(* IEC 61131-3 sources: stdmachine/plc/src/04_Objects, 21 files *)

(* ---- FB_AnalogInput.st ---- *)
// Entrée analogique, type 3 (docs/03 § 3.3)
FUNCTION_BLOCK FB_AnalogInput EXTENDS FB_ObjectBase
VAR
    _aSamples : ARRAY[1..100] OF LREAL;
    _nSamples : INT;
    _nNext : INT := 1;
    _fValue : LREAL;                // valeur filtrée, en unité
    _bLowActive : BOOL;
    _bHighActive : BOOL;
END_VAR

METHOD PROTECTED _OnConfigure : BOOL
_nSamples := 0;
_nNext := 1;
_OnConfigure := F_SignalValid(_refCfg.aSignal[1], E_SignalKind.AI) AND _refCfg.aParam[2] <> _refCfg.aParam[1];
END_METHOD

METHOD PROTECTED _OnStart : E_ActStatus
VAR_INPUT
    nAction : UINT;
END_VAR
CASE nAction OF
    GVL_Catalog.AnalogInput_Lire:
        _SetResult(1, _fValue);
        _OnStart := E_ActStatus.Done;
    GVL_Catalog.AnalogInput_AttendreSeuil:
        _OnStart := _OnCycle(nAction);
    GVL_Catalog.AnalogInput_VerifierPlage:
        _SetResult(1, _fValue);
        IF _fValue < _ParamReal(1, -1.0E38) THEN
            _SetJudgement(2, E_Judgement.Low);
        ELSIF _fValue > _ParamReal(2, 1.0E38) THEN
            _SetJudgement(2, E_Judgement.High);
        ELSE
            _SetJudgement(2, E_Judgement.Ok);
        END_IF
        _OnStart := E_ActStatus.Done;
ELSE
    _OnStart := E_ActStatus.Error;
END_CASE
END_METHOD

METHOD PROTECTED _OnCycle : E_ActStatus
VAR_INPUT
    nAction : UINT;
END_VAR
VAR
    bReached : BOOL;
END_VAR
IF _ParamReal(2, 0.0) = 0.0 THEN
    bReached := _fValue >= _ParamReal(1, 0.0);      // au-dessus
ELSE
    bReached := _fValue <= _ParamReal(1, 0.0);      // en dessous
END_IF
IF bReached THEN
    _SetResult(1, _fValue);
    _OnCycle := E_ActStatus.Done;
ELSE
    _OnCycle := E_ActStatus.Busy;
END_IF
END_METHOD

METHOD PROTECTED _ReadHw
_Filter(_Scale(INT_TO_LREAL(F_ReadAI(_refCfg.aSignal[1]))));
END_METHOD

METHOD PROTECTED _Simulate
IF _Forced(1) THEN _Filter(_ForcedValue(1)); END_IF        // valeur forcée en unité
END_METHOD

METHOD PRIVATE _Scale : LREAL
VAR_INPUT
    fRaw : LREAL;
END_VAR
_Scale := _refCfg.aParam[3] + (fRaw - _refCfg.aParam[1]) * (_refCfg.aParam[4] - _refCfg.aParam[3]) / (_refCfg.aParam[2] - _refCfg.aParam[1]);
END_METHOD

METHOD PRIVATE _Filter
VAR_INPUT
    fUnit : LREAL;
END_VAR
VAR
    nWin : INT;
    i : INT;
    fSum : LREAL;
END_VAR
nWin := LIMIT(1, LREAL_TO_INT(_refCfg.aParam[6]), 100);
_aSamples[_nNext] := fUnit;
_nNext := _nNext MOD nWin + 1;
_nSamples := MIN(_nSamples + 1, nWin);
fSum := 0;
FOR i := 1 TO _nSamples DO fSum := fSum + _aSamples[i]; END_FOR
_fValue := fSum / INT_TO_LREAL(_nSamples);
END_METHOD

// Seuils d'alarme : avertissements surveillés en continu, sans mettre l'objet en erreur
METHOD PROTECTED _Monitor
IF _ipAlarms = 0 THEN RETURN; END_IF
IF _fValue < _refCfg.aParam[7] AND NOT _bLowActive THEN
    _ipAlarms.Raise(_stInfo.nGlobalId, GVL_Catalog.AnalogInput_Err100, 0, E_Severity.Warning);
    _bLowActive := TRUE;
ELSIF _fValue >= _refCfg.aParam[7] AND _bLowActive THEN
    _ipAlarms.Clear(_stInfo.nGlobalId, GVL_Catalog.AnalogInput_Err100);
    _bLowActive := FALSE;
END_IF
IF _fValue > _refCfg.aParam[8] AND NOT _bHighActive THEN
    _ipAlarms.Raise(_stInfo.nGlobalId, GVL_Catalog.AnalogInput_Err101, 0, E_Severity.Warning);
    _bHighActive := TRUE;
ELSIF _fValue <= _refCfg.aParam[8] AND _bHighActive THEN
    _ipAlarms.Clear(_stInfo.nGlobalId, GVL_Catalog.AnalogInput_Err101);
    _bHighActive := FALSE;
END_IF
END_METHOD

METHOD PROTECTED _Publish
_stStatus.aValue[1] := _fValue;
END_METHOD

PROPERTY Value : LREAL
GET
Value := _fValue;
END_GET
END_PROPERTY
END_FUNCTION_BLOCK

(* ---- FB_AnalogOutput.st ---- *)
// Sortie analogique, type 4 (docs/03 § 3.4)
FUNCTION_BLOCK FB_AnalogOutput EXTENDS FB_ObjectBase
VAR
    _fValue : LREAL;                // valeur commandée, en unité
    _fStart : LREAL;
    _fTarget : LREAL;
    _fRampMs : LREAL;
    _fElapsed : LREAL;
END_VAR

METHOD PROTECTED _OnConfigure : BOOL
_OnConfigure := F_SignalValid(_refCfg.aSignal[1], E_SignalKind.AO) AND _refCfg.aParam[4] <> _refCfg.aParam[3];
END_METHOD

METHOD PROTECTED _DefaultTimeoutMs : UDINT
VAR_INPUT
    nAction : UINT;
END_VAR
IF nAction = GVL_Catalog.AnalogOutput_EcrireAvecRampe THEN
    _DefaultTimeoutMs := LREAL_TO_UDINT(MAX(_ParamReal(2, 0.0), 0.0)) + 1000;
ELSE
    _DefaultTimeoutMs := 0;
END_IF
END_METHOD

METHOD PROTECTED _OnStart : E_ActStatus
VAR_INPUT
    nAction : UINT;
END_VAR
_fStart := _fValue;
_fElapsed := 0;
CASE nAction OF
    GVL_Catalog.AnalogOutput_Ecrire:
        _fTarget := _Limit(_ParamReal(1, _fValue));
        _fRampMs := 0;
    GVL_Catalog.AnalogOutput_EcrireAvecRampe:
        _fTarget := _Limit(_ParamReal(1, _fValue));
        _fRampMs := MAX(_ParamReal(2, 0.0), 0.0);
    GVL_Catalog.AnalogOutput_ValeurSure:
        _fTarget := _Limit(_refCfg.aParam[8]);
        _fRampMs := 0;
ELSE
    _OnStart := E_ActStatus.Error;
    RETURN;
END_CASE
_OnStart := _OnCycle(nAction);
END_METHOD

METHOD PROTECTED _OnCycle : E_ActStatus
VAR_INPUT
    nAction : UINT;
END_VAR
VAR
    fNext : LREAL;
    fMaxStep : LREAL;
END_VAR
_fElapsed := _fElapsed + F_CycleMs();
IF _fRampMs > 0 THEN
    fNext := _fStart + (_fTarget - _fStart) * MIN(1.0, _fElapsed / _fRampMs);
ELSE
    fNext := _fTarget;
END_IF
// Variation maximale P9 (unité/s), 0 = illimitée
IF _refCfg.aParam[9] > 0 THEN
    fMaxStep := _refCfg.aParam[9] * F_CycleMs() / 1000.0;
    fNext := LIMIT(_fValue - fMaxStep, fNext, _fValue + fMaxStep);
END_IF
_fValue := fNext;
IF ABS(_fValue - _fTarget) < 1.0E-9 THEN _OnCycle := E_ActStatus.Done; ELSE _OnCycle := E_ActStatus.Busy; END_IF
END_METHOD

METHOD PRIVATE _Limit : LREAL
VAR_INPUT
    fValue : LREAL;
END_VAR
_Limit := LIMIT(_refCfg.aParam[6], fValue, _refCfg.aParam[7]);
END_METHOD

METHOD PROTECTED _SafeState
_fValue := _Limit(_refCfg.aParam[8]);
END_METHOD

METHOD PROTECTED _WriteHw
VAR
    fRaw : LREAL;
END_VAR
fRaw := _refCfg.aParam[1] + (_fValue - _refCfg.aParam[3]) * (_refCfg.aParam[2] - _refCfg.aParam[1]) / (_refCfg.aParam[4] - _refCfg.aParam[3]);
F_WriteAO(_refCfg.aSignal[1], LREAL_TO_INT(LIMIT(-32768.0, fRaw, 32767.0)));
END_METHOD

METHOD PROTECTED _Publish
_stStatus.aValue[1] := _fValue;
END_METHOD
END_FUNCTION_BLOCK

(* ---- FB_Axis.st ---- *)
// Axe linéaire (type 11) et axe rotatif (type 12), docs/03 § 4.2 et docs/04 § 12.
// Matériel : D = n° de l'axe dans GVL_Hw.aAxis (pointeur donné par GVL_IoRef). Blocs Tc2_MC2.
// L'override effectif est appliqué par MC_Power.Override : il ralentit le mouvement en cours sans le relancer.
FUNCTION_BLOCK FB_Axis EXTENDS FB_ObjectBase
VAR
    _pAxis : POINTER TO AXIS_REF;
    _bRotary : BOOL;
    _fbPower : MC_Power;
    _fbReset : MC_Reset;
    _fbHome : MC_Home;
    _fbMoveAbs : MC_MoveAbsolute;
    _fbMoveMod : MC_MoveModulo;
    _fbMoveRel : MC_MoveRelative;
    _fbHalt : MC_Halt;
    _fbStop : MC_Stop;
    _fbJog : MC_Jog;
    _bEnable : BOOL;                // alimentation demandée
    _bPowered : BOOL;
    _bWasPowered : BOOL;
    _bHomed : BOOL;
    _fActPos : LREAL;
    _fActVel : LREAL;
    _fTarget : LREAL;
    _fStartPos : LREAL;
    _fVelo : LREAL;
    _fAcc : LREAL;
    _fDec : LREAL;
    _nDirection : INT;              // rotatif : 0 plus court, 1 positif, 2 négatif
    _bExecute : BOOL;               // front de commande de l'action en cours
    _bStopping : BOOL;              // Abort : arrêt en cours
    _fOverride : LREAL := 100.0;
    // Simulation : profil trapézoïdal
    _fSimPos : LREAL;
    _fSimVel : LREAL;
    _fSimInitMs : LREAL;
    _nJogDir : INT;                 // +1, -1, 0
END_VAR

METHOD PROTECTED _OnConfigure : BOOL
_bRotary := _refCfg.nType = GVL_Catalog.Type_RotaryAxis;
_pAxis := F_AxisRef(_refCfg.nDevice);
_bEnable := FALSE;
_bHomed := FALSE;
_fSimVel := 0;
_OnConfigure := _pAxis <> 0 OR _IsSimulated();
END_METHOD

METHOD PROTECTED _NeedsInit : BOOL
_NeedsInit := TRUE;
END_METHOD

METHOD PROTECTED _IsAllowedNotInit : BOOL
VAR_INPUT
    nAction : UINT;
END_VAR
_IsAllowedNotInit := nAction = GVL_Catalog.LinearAxis_PowerOn OR nAction = GVL_Catalog.LinearAxis_PowerOff
                     OR nAction = GVL_Catalog.LinearAxis_Init OR nAction = GVL_Catalog.LinearAxis_AcquitterErreur
                     OR nAction = GVL_Catalog.LinearAxis_LirePosition
                     OR nAction = GVL_Catalog.LinearAxis_JogPlus OR nAction = GVL_Catalog.LinearAxis_JogMoins;
END_METHOD

METHOD PROTECTED _ManualOverride : LREAL
_ManualOverride := LIMIT(0.0, _refCfg.aParam[12], 100.0);
END_METHOD

METHOD PROTECTED _DefaultTimeoutMs : UDINT
VAR_INPUT
    nAction : UINT;
END_VAR
VAR
    fDist : LREAL;
END_VAR
// Move absolu et relatif : 2 × (distance ÷ vitesse + vitesse ÷ accélération) × 1000 + 1000 ms, à 100 %
IF nAction = GVL_Catalog.LinearAxis_MoveAbsolu OR nAction = GVL_Catalog.LinearAxis_MoveRelatif THEN
    IF nAction = GVL_Catalog.LinearAxis_MoveAbsolu THEN fDist := ABS(_TargetOf() - _fActPos); ELSE fDist := ABS(_ParamReal(1, 0.0)); END_IF
    _Kinematics();
    IF _fVelo > 0 AND _fAcc > 0 THEN
        _DefaultTimeoutMs := LREAL_TO_UDINT(2.0 * (fDist / _fVelo + _fVelo / _fAcc) * 1000.0 + 1000.0);
    ELSE
        _DefaultTimeoutMs := 30000;
    END_IF
ELSE
    _DefaultTimeoutMs := SUPER^._DefaultTimeoutMs(nAction);
END_IF
END_METHOD

METHOD PRIVATE _TargetOf : LREAL
// Une position nommée : composante P13 (X, Y, Z) ou C pour un rotatif, plus le décalage (hauteur d'approche)
IF _stParams.aKind[1] = E_ParamKind.Position THEN
    IF _bRotary THEN
        _TargetOf := _stParams.stPos.fC;
    ELSE
        CASE LREAL_TO_INT(_refCfg.aParam[13]) OF
            1: _TargetOf := _stParams.stPos.fY;
            2: _TargetOf := _stParams.stPos.fZ;
        ELSE
            _TargetOf := _stParams.stPos.fX;
        END_CASE
    END_IF
    _TargetOf := _TargetOf + _stParams.aReal[1];
ELSE
    _TargetOf := _stParams.aReal[1];
END_IF
END_METHOD

METHOD PRIVATE _Kinematics
VAR
    fAccPct : LREAL;
END_VAR
_fVelo := MAX(_refCfg.aParam[1], 0.001) * F_ParamSpeed(_stParams, 2, _refCfg, 2) / 100.0;
fAccPct := LIMIT(1.0, _ParamReal(3, 100.0), 100.0);
IF _stParams.aKind[3] = E_ParamKind.Unused THEN fAccPct := 100.0; END_IF
_fAcc := MAX(_refCfg.aParam[2], 0.001) * fAccPct / 100.0;
_fDec := MAX(_refCfg.aParam[3], 0.001) * fAccPct / 100.0;
END_METHOD

METHOD PROTECTED _OnStart : E_ActStatus
VAR_INPUT
    nAction : UINT;
END_VAR
_bExecute := FALSE;
_bStopping := FALSE;
_fStartPos := _fActPos;
CASE nAction OF
    GVL_Catalog.LinearAxis_PowerOn:
        _bEnable := TRUE;
        _OnStart := E_ActStatus.Busy;
    GVL_Catalog.LinearAxis_PowerOff:
        _bEnable := FALSE;
        _OnStart := E_ActStatus.Busy;
    GVL_Catalog.LinearAxis_Init:
        IF NOT _bPowered THEN _Fail(GVL_Catalog.LinearAxis_Err105, 0); _OnStart := E_ActStatus.Error; RETURN; END_IF
        _bHomed := FALSE;
        _bInitialized := FALSE;
        _fSimInitMs := 0;
        _OnStart := E_ActStatus.Busy;
    GVL_Catalog.LinearAxis_MoveAbsolu, GVL_Catalog.LinearAxis_MoveRelatif:
        IF NOT _bPowered THEN _Fail(GVL_Catalog.LinearAxis_Err105, 0); _OnStart := E_ActStatus.Error; RETURN; END_IF
        IF NOT _bHomed THEN _Fail(GVL_Catalog.LinearAxis_Err100, 0); _OnStart := E_ActStatus.Error; RETURN; END_IF
        IF nAction = GVL_Catalog.LinearAxis_MoveAbsolu THEN
            _fTarget := _TargetOf();
            _nDirection := LREAL_TO_INT(_ParamReal(4, _refCfg.aParam[14]));
        ELSE
            _fTarget := _fActPos + _ParamReal(1, 0.0);
        END_IF
        IF _refCfg.aParam[7] = 1 AND (_fTarget < _refCfg.aParam[5] OR _fTarget > _refCfg.aParam[6]) THEN
            _Fail(GVL_Catalog.LinearAxis_Err101, 0);
            _OnStart := E_ActStatus.Error;
            RETURN;
        END_IF
        _Kinematics();
        _OnStart := E_ActStatus.Busy;
    GVL_Catalog.LinearAxis_Stop:
        _OnStart := E_ActStatus.Busy;
    GVL_Catalog.LinearAxis_AcquitterErreur:
        _OnStart := E_ActStatus.Busy;
    GVL_Catalog.LinearAxis_LirePosition:
        _SetResult(1, _fActPos);
        _OnStart := E_ActStatus.Done;
    GVL_Catalog.LinearAxis_JogPlus, GVL_Catalog.LinearAxis_JogMoins:
        IF NOT _bPowered THEN _Fail(GVL_Catalog.LinearAxis_Err105, 0); _OnStart := E_ActStatus.Error; RETURN; END_IF
        _fVelo := MAX(_refCfg.aParam[1], 0.001) * F_ParamSpeed(_stParams, 1, _refCfg, 1) / 100.0;
        IF NOT _bHomed THEN _fVelo := MAX(_refCfg.aParam[1], 0.001) * F_ParamSpeed(_stParams, 0, _refCfg, 1) / 100.0; END_IF   // V1 imposée
        _fAcc := MAX(_refCfg.aParam[2], 0.001);
        _fDec := MAX(_refCfg.aParam[3], 0.001);
        _nJogDir := SEL(nAction = GVL_Catalog.LinearAxis_JogPlus, -1, 1);
        _OnStart := E_ActStatus.Busy;       // le jog dure jusqu'à Abort (canal manuel, docs/05 § 7)
ELSE
    _OnStart := E_ActStatus.Error;
END_CASE
END_METHOD

METHOD PROTECTED _OnCycle : E_ActStatus
VAR_INPUT
    nAction : UINT;
END_VAR
_OnCycle := E_ActStatus.Busy;
CASE nAction OF
    GVL_Catalog.LinearAxis_PowerOn:
        IF _bPowered THEN _OnCycle := E_ActStatus.Done; END_IF
    GVL_Catalog.LinearAxis_PowerOff:
        IF NOT _bPowered THEN _OnCycle := E_ActStatus.Done; END_IF
    GVL_Catalog.LinearAxis_Init:
        IF _IsSimulated() THEN
            _fSimInitMs := _fSimInitMs + F_CycleMs();
            IF _fSimInitMs >= 1500.0 THEN
                _fSimPos := _refCfg.aParam[8];
                _fSimVel := 0;
                _bHomed := TRUE;
            END_IF
        ELSE
            _bExecute := TRUE;
            IF _fbHome.Done THEN _bHomed := TRUE; END_IF
            IF _fbHome.Error THEN _Fail(GVL_Catalog.LinearAxis_Err102, _fbHome.ErrorID); _OnCycle := E_ActStatus.Error; RETURN; END_IF
        END_IF
        IF _bHomed THEN
            _bInitialized := TRUE;
            _bExecute := FALSE;
            _OnCycle := E_ActStatus.Done;
        END_IF
    GVL_Catalog.LinearAxis_MoveAbsolu, GVL_Catalog.LinearAxis_MoveRelatif:
        IF _IsSimulated() THEN
            IF ABS(_fSimPos - _fTarget) <= MAX(_refCfg.aParam[4], 1.0E-6) AND ABS(_fSimVel) < 1.0E-6 THEN _OnCycle := E_ActStatus.Done; END_IF
        ELSE
            _bExecute := TRUE;
            IF _fbMoveAbs.Done OR _fbMoveRel.Done OR _fbMoveMod.Done THEN _OnCycle := E_ActStatus.Done; END_IF
            IF _fbMoveAbs.Error OR _fbMoveRel.Error OR _fbMoveMod.Error THEN
                _Fail(GVL_Catalog.LinearAxis_Err102, _fbMoveAbs.ErrorID OR _fbMoveRel.ErrorID OR _fbMoveMod.ErrorID);
                _OnCycle := E_ActStatus.Error;
                RETURN;
            END_IF
        END_IF
        IF _OnCycle = E_ActStatus.Done THEN
            _bExecute := FALSE;
            _SetResult(1, _fActPos);
        END_IF
    GVL_Catalog.LinearAxis_Stop:
        IF _IsSimulated() THEN
            IF ABS(_fSimVel) < 1.0E-6 THEN _OnCycle := E_ActStatus.Done; END_IF
        ELSE
            _bExecute := TRUE;
            IF _fbHalt.Done THEN _bExecute := FALSE; _OnCycle := E_ActStatus.Done; END_IF
        END_IF
    GVL_Catalog.LinearAxis_AcquitterErreur:
        IF _IsSimulated() THEN
            _OnCycle := E_ActStatus.Done;
        ELSE
            _bExecute := TRUE;
            IF _fbReset.Done OR _fbReset.Error THEN _bExecute := FALSE; _OnCycle := E_ActStatus.Done; END_IF
        END_IF
    GVL_Catalog.LinearAxis_JogPlus, GVL_Catalog.LinearAxis_JogMoins:
        ;                               // jusqu'à Abort
END_CASE
_CallMotion();
END_METHOD

METHOD PROTECTED _OnAbort
VAR_INPUT
    nAction : UINT;
END_VAR
// Arrêt avec la décélération maximale, puis P11 (0 alimentation maintenue, 1 coupée)
_bExecute := FALSE;
_nJogDir := 0;
_bStopping := TRUE;
END_METHOD

METHOD PROTECTED _SafeState
IF _refCfg.aParam[11] = 1 THEN _bEnable := FALSE; END_IF
END_METHOD

METHOD PROTECTED _OnAck : BOOL
IF _IsSimulated() OR _pAxis = 0 THEN
    _OnAck := TRUE;
    RETURN;
END_IF
_fbReset(Axis := _pAxis^, Execute := TRUE);
IF _fbReset.Done OR _fbReset.Error THEN
    _fbReset(Axis := _pAxis^, Execute := FALSE);
    _OnAck := TRUE;
END_IF
END_METHOD

METHOD PROTECTED _ApplyOverride
VAR_INPUT
    fPercent : LREAL;
END_VAR
_fOverride := LIMIT(0.0, fPercent, 100.0);
END_METHOD

METHOD PROTECTED _ReadHw
IF _pAxis = 0 THEN RETURN; END_IF
_pAxis^.ReadStatus();
_fActPos := _pAxis^.NcToPlc.ActPos;
_fActVel := _pAxis^.NcToPlc.ActVelo;
_bHomed := _bHomed OR _pAxis^.Status.Homed;
_fbPower(Axis := _pAxis^, Enable := _bEnable, Enable_Positive := _bEnable, Enable_Negative := _bEnable, Override := _fOverride);
_bPowered := _fbPower.Status;
IF NOT _bExecute AND _eState <> E_ObjState.Busy THEN _CallMotion(); END_IF    // remet les Execute à FALSE
END_METHOD

METHOD PRIVATE _CallMotion
VAR
    bAbs : BOOL;
    bRel : BOOL;
    bMod : BOOL;
    eDir : MC_Direction;
END_VAR
IF _IsSimulated() OR _pAxis = 0 THEN RETURN; END_IF
bAbs := _bExecute AND _nAction = GVL_Catalog.LinearAxis_MoveAbsolu AND NOT (_bRotary AND _refCfg.aParam[7] = 0);
bMod := _bExecute AND _nAction = GVL_Catalog.LinearAxis_MoveAbsolu AND _bRotary AND _refCfg.aParam[7] = 0;
bRel := _bExecute AND _nAction = GVL_Catalog.LinearAxis_MoveRelatif;
CASE _nDirection OF
    1: eDir := MC_Positive_Direction;
    2: eDir := MC_Negative_Direction;
ELSE
    eDir := MC_Shortest_Way;
END_CASE
_fbHome(Axis := _pAxis^, Execute := _bExecute AND _nAction = GVL_Catalog.LinearAxis_Init, Position := _refCfg.aParam[8],
        HomingMode := SEL(LREAL_TO_INT(_refCfg.aParam[9]) = 3, MC_DefaultHoming, MC_Direct));
_fbMoveAbs(Axis := _pAxis^, Execute := bAbs, Position := _fTarget, Velocity := _fVelo, Acceleration := _fAcc, Deceleration := _fDec);
_fbMoveMod(Axis := _pAxis^, Execute := bMod, Position := _fTarget, Velocity := _fVelo, Acceleration := _fAcc, Deceleration := _fDec, Direction := eDir);
_fbMoveRel(Axis := _pAxis^, Execute := bRel, Distance := _fTarget - _fStartPos, Velocity := _fVelo, Acceleration := _fAcc, Deceleration := _fDec);
_fbHalt(Axis := _pAxis^, Execute := _bExecute AND _nAction = GVL_Catalog.LinearAxis_Stop);
_fbReset(Axis := _pAxis^, Execute := _bExecute AND _nAction = GVL_Catalog.LinearAxis_AcquitterErreur);
_fbJog(Axis := _pAxis^, JogForward := _nJogDir > 0, JogBackwards := _nJogDir < 0, Mode := MC_JOGMODE_CONTINOUS,
       Velocity := _fVelo, Acceleration := _fAcc, Deceleration := _fDec);
_fbStop(Axis := _pAxis^, Execute := _bStopping);
IF _bStopping AND (_fbStop.Done OR _fbStop.Error) THEN
    _bStopping := FALSE;
    _fbStop(Axis := _pAxis^, Execute := FALSE);
END_IF
END_METHOD

METHOD PROTECTED _Monitor
IF _IsSimulated() OR _pAxis = 0 THEN
    _bWasPowered := _bPowered;
    RETURN;
END_IF
IF _pAxis^.Status.Error AND _eState <> E_ObjState.Error THEN
    IF _pAxis^.Status.ErrorID = 16#4550 OR _pAxis^.Status.ErrorID = 16#4551 THEN
        _Fail(GVL_Catalog.LinearAxis_Err103, _pAxis^.Status.ErrorID);      // erreur de suivi
    ELSE
        _Fail(GVL_Catalog.LinearAxis_Err102, _pAxis^.Status.ErrorID);      // erreur du drive (sous-code NC)
    END_IF
ELSIF _bWasPowered AND NOT _bPowered AND _bEnable AND _eState <> E_ObjState.Error THEN
    _Fail(GVL_Catalog.LinearAxis_Err104, 0);                                 // perte d'alimentation
END_IF
_bWasPowered := _bPowered;
END_METHOD

METHOD PROTECTED _Simulate
VAR
    fDt : LREAL;
    fVmax : LREAL;
    fDist : LREAL;
    fBrake : LREAL;
    fDir : LREAL;
END_VAR
fDt := F_CycleMs() / 1000.0;
_bPowered := _bEnable;
fVmax := _fVelo * _fOverride / 100.0;
IF _bStopping THEN
    // arrêt avec la décélération maximale
    IF _fSimVel > 0 THEN _fSimVel := MAX(0.0, _fSimVel - _refCfg.aParam[3] * fDt); ELSE _fSimVel := MIN(0.0, _fSimVel + _refCfg.aParam[3] * fDt); END_IF
    IF ABS(_fSimVel) < 1.0E-9 THEN _bStopping := FALSE; END_IF
ELSIF _eState = E_ObjState.Busy AND (_nAction = GVL_Catalog.LinearAxis_JogPlus OR _nAction = GVL_Catalog.LinearAxis_JogMoins) THEN
    _fSimVel := LIMIT(-fVmax, _fSimVel + INT_TO_LREAL(_nJogDir) * _fAcc * fDt, fVmax);
ELSIF _eState = E_ObjState.Busy AND (_nAction = GVL_Catalog.LinearAxis_MoveAbsolu OR _nAction = GVL_Catalog.LinearAxis_MoveRelatif) THEN
    fDist := _fTarget - _fSimPos;
    fDir := SEL(fDist >= 0, -1.0, 1.0);
    fBrake := _fSimVel * _fSimVel / (2.0 * MAX(_fDec, 0.001));
    IF ABS(fDist) <= fBrake THEN
        _fSimVel := _fSimVel - fDir * _fDec * fDt;          // décélération
        IF fDir * _fSimVel < 0 THEN _fSimVel := 0; END_IF
    ELSE
        _fSimVel := LIMIT(-fVmax, _fSimVel + fDir * _fAcc * fDt, fVmax);
    END_IF
    IF ABS(fDist) <= ABS(_fSimVel * fDt) OR (ABS(_fSimVel) < 1.0E-9 AND ABS(fDist) <= MAX(_refCfg.aParam[4], 1.0E-6)) THEN
        _fSimPos := _fTarget;
        _fSimVel := 0;
    END_IF
ELSIF _eState = E_ObjState.Busy AND _nAction = GVL_Catalog.LinearAxis_Stop THEN
    IF _fSimVel > 0 THEN _fSimVel := MAX(0.0, _fSimVel - _fDec * fDt); ELSE _fSimVel := MIN(0.0, _fSimVel + _fDec * fDt); END_IF
ELSE
    _fSimVel := 0;
END_IF
_fSimPos := _fSimPos + _fSimVel * fDt;
_fActPos := _fSimPos;
_fActVel := _fSimVel;
END_METHOD

METHOD PROTECTED _Publish
_stStatus.aValue[1] := _fActPos;
_stStatus.aValue[2] := _fActVel;
_stStatus.aValue[3] := BOOL_TO_LREAL(_bPowered);
_stStatus.aValue[4] := BOOL_TO_LREAL(_bHomed);
IF _eState = E_ObjState.Busy AND ABS(_fTarget - _fStartPos) > 1.0E-9
   AND (_nAction = GVL_Catalog.LinearAxis_MoveAbsolu OR _nAction = GVL_Catalog.LinearAxis_MoveRelatif) THEN
    _stStatus.fProgress := LREAL_TO_REAL(LIMIT(0.0, ABS(_fActPos - _fStartPos) / ABS(_fTarget - _fStartPos), 1.0));
END_IF
END_METHOD

PROPERTY ActualPosition : LREAL
GET
ActualPosition := _fActPos;
END_GET
END_PROPERTY
END_FUNCTION_BLOCK

(* ---- FB_Beacon.st ---- *)
// Balise, type 50 (docs/03 § 8.1) : pilotée par le séquenceur ; actions de test en manuel seulement
FUNCTION_BLOCK FB_Beacon EXTENDS FB_ObjectBase IMPLEMENTS I_Beacon
VAR
    _nPattern : UINT;
    _bBuzzerReq : BOOL;
    _fBlink : LREAL;
    _bPhase : BOOL;
    _nTestColor : INT := -1;        // test manuel : 0 rouge, 1 orange, 2 vert, 3 bleu, 4 buzzer
    _fTestMs : LREAL;
    _fBuzzMs : LREAL;               // durée de buzzer demandée (0 = jusqu'à acquittement)
    _fBuzzElapsed : LREAL;
    _aOut : ARRAY[1..5] OF BOOL;    // rouge, orange, vert, bleu, buzzer
END_VAR

METHOD SetPattern
VAR_INPUT
    nPattern : UINT;
    bBuzzer : BOOL;
END_VAR
IF bBuzzer AND NOT _bBuzzerReq THEN _fBuzzElapsed := 0; END_IF
_nPattern := nPattern;
_bBuzzerReq := bBuzzer;
END_METHOD

METHOD PROTECTED _OnStart : E_ActStatus
VAR_INPUT
    nAction : UINT;
END_VAR
_fBuzzElapsed := 0;
CASE nAction OF
    GVL_Catalog.Beacon_Tester:
        _nTestColor := LIMIT(0, LREAL_TO_INT(_ParamReal(1, 0.0)), 4);
        _fTestMs := MAX(_ParamReal(2, 2000.0), 100.0);
        _OnStart := E_ActStatus.Busy;
    GVL_Catalog.Beacon_Buzzer:
        _nTestColor := 4;
        _fTestMs := MAX(_ParamReal(1, 1000.0), 100.0);
        _OnStart := E_ActStatus.Busy;
ELSE
    _OnStart := E_ActStatus.Error;
END_CASE
END_METHOD

METHOD PROTECTED _OnCycle : E_ActStatus
VAR_INPUT
    nAction : UINT;
END_VAR
IF _fElapsedMs >= _fTestMs THEN
    _nTestColor := -1;
    _OnCycle := E_ActStatus.Done;
ELSE
    _OnCycle := E_ActStatus.Busy;
END_IF
END_METHOD

METHOD PROTECTED _OnAbort
VAR_INPUT
    nAction : UINT;
END_VAR
_nTestColor := -1;
END_METHOD

METHOD PROTECTED _Monitor
VAR
    fPeriod : LREAL;
    i : INT;
END_VAR
fPeriod := MAX(_refCfg.aParam[1], 100.0);
_fBlink := _fBlink + F_CycleMs();
IF _fBlink >= fPeriod / 2.0 THEN
    _fBlink := 0;
    _bPhase := NOT _bPhase;
END_IF
FOR i := 1 TO 5 DO _aOut[i] := FALSE; END_FOR
IF _nTestColor >= 0 THEN
    _aOut[_nTestColor + 1] := TRUE;
    RETURN;
END_IF
_aOut[1] := (_nPattern AND GVL_BeaconBits.RED) <> 0 OR ((_nPattern AND GVL_BeaconBits.RED_BLINK) <> 0 AND _bPhase);
_aOut[2] := (_nPattern AND GVL_BeaconBits.ORANGE) <> 0 OR ((_nPattern AND GVL_BeaconBits.ORANGE_BLINK) <> 0 AND _bPhase);
_aOut[3] := (_nPattern AND GVL_BeaconBits.GREEN) <> 0 OR ((_nPattern AND GVL_BeaconBits.GREEN_BLINK) <> 0 AND _bPhase);
_aOut[4] := (_nPattern AND GVL_BeaconBits.BLUE) <> 0 OR ((_nPattern AND GVL_BeaconBits.BLUE_BLINK) <> 0 AND _bPhase);
IF _bBuzzerReq THEN
    _fBuzzElapsed := _fBuzzElapsed + F_CycleMs();
    _aOut[5] := _refCfg.aParam[2] <= 0 OR _fBuzzElapsed < _refCfg.aParam[2];
END_IF
END_METHOD

METHOD PROTECTED _WriteHw
VAR
    i : USINT;
END_VAR
FOR i := 1 TO 5 DO F_WriteDO(_refCfg.aSignal[i], _aOut[i]); END_FOR
END_METHOD

METHOD PROTECTED _Publish
VAR
    i : INT;
    nBits : DWORD;
END_VAR
FOR i := 1 TO 5 DO
    IF _aOut[i] THEN nBits := nBits OR SHL(DWORD#1, i - 1); END_IF
END_FOR
_stStatus.aValue[1] := DWORD_TO_LREAL(nBits);
END_METHOD
END_FUNCTION_BLOCK

(* ---- FB_Counter.st ---- *)
// Compteur, type 53 (docs/03 § 8.4)
FUNCTION_BLOCK FB_Counter EXTENDS FB_ObjectBase IMPLEMENTS I_OrderAware
VAR
    _bStarted : BOOL;               // faux au démarrage du PLC (P4 = 0 : la valeur repart de P1)
END_VAR
VAR PERSISTENT
    _fValue : LREAL;
END_VAR

METHOD PROTECTED _OnConfigure : BOOL
IF _bNewObject THEN _fValue := _refCfg.aParam[1]; END_IF
_OnConfigure := TRUE;
END_METHOD

METHOD PROTECTED _OnStart : E_ActStatus
VAR_INPUT
    nAction : UINT;
END_VAR
CASE nAction OF
    GVL_Catalog.Counter_Incrementer:
        _fValue := _fValue + _ParamReal(1, 1.0);
        _SetResult(1, _fValue);
        IF _refCfg.aParam[2] > 0 AND _fValue > _refCfg.aParam[2] THEN
            _Fail(GVL_Catalog.Counter_Err100, LREAL_TO_UDINT(_fValue));
            _OnStart := E_ActStatus.Error;
            RETURN;
        END_IF
    GVL_Catalog.Counter_Lire:
        _SetResult(1, _fValue);
    GVL_Catalog.Counter_RemettreAZero:
        _fValue := _refCfg.aParam[1];
    GVL_Catalog.Counter_Comparer:
        _SetResult(1, BOOL_TO_LREAL(_fValue >= _ParamReal(1, 0.0)));
ELSE
    _OnStart := E_ActStatus.Error;
    RETURN;
END_CASE
_OnStart := E_ActStatus.Done;
END_METHOD

// Remise à zéro au changement d'OF (P3), appelée par le séquenceur général
METHOD OnOrderChange
IF _refCfg.aParam[3] = 1 THEN _fValue := _refCfg.aParam[1]; END_IF
END_METHOD

METHOD PROTECTED _Monitor
IF NOT _bStarted THEN
    _bStarted := TRUE;
    IF _refCfg.aParam[4] = 0 THEN _fValue := _refCfg.aParam[1]; END_IF
END_IF
END_METHOD

METHOD PROTECTED _Publish
_stStatus.aValue[1] := _fValue;
END_METHOD
END_FUNCTION_BLOCK

(* ---- FB_Cylinder.st ---- *)
// Vérin, type 10 (docs/03 § 4.1, exemple complet de docs/04 § 11)
FUNCTION_BLOCK FB_Cylinder EXTENDS FB_ObjectBase
VAR
    _bBistable : BOOL;
    _tSettleMs : LREAL;
    _tNoSensorMs : LREAL;
    _eSafe : USINT;                 // 0 Repos, 1 Travail, 2 Maintien
    _bCmdWork : BOOL;               // sortie travail commandée
    _bAtWork : BOOL;                // capteurs (lus ou simulés)
    _bAtRest : BOOL;
    _bHasWorkSensor : BOOL;
    _bHasRestSensor : BOOL;
    _fSettle : LREAL;
    _fMove : LREAL;
    _fSimPos : LREAL;               // simulation : 0 = repos, 1 = travail
    _nReached : USINT;              // 0 aucune, 1 repos, 2 travail : dernière position atteinte par une action
END_VAR

METHOD PROTECTED _OnConfigure : BOOL
_bBistable := _refCfg.aParam[1] = 1;
_tSettleMs := LIMIT(0.0, _refCfg.aParam[2], 5000.0);
_tNoSensorMs := MAX(_refCfg.aParam[3], 10.0);
_eSafe := LREAL_TO_USINT(_refCfg.aParam[4]);
_bHasWorkSensor := F_SignalValid(_refCfg.aSignal[3], E_SignalKind.DI);
_bHasRestSensor := F_SignalValid(_refCfg.aSignal[4], E_SignalKind.DI);
_nReached := 0;
_OnConfigure := F_SignalValid(_refCfg.aSignal[1], E_SignalKind.DO)
                AND (NOT _bBistable OR F_SignalValid(_refCfg.aSignal[2], E_SignalKind.DO));
END_METHOD

METHOD PROTECTED _DefaultTimeoutMs : UDINT
VAR_INPUT
    nAction : UINT;
END_VAR
_DefaultTimeoutMs := SEL(_bHasWorkSensor OR _bHasRestSensor, LREAL_TO_UDINT(_tNoSensorMs) + 500, 2000);
END_METHOD

METHOD PROTECTED _OnStart : E_ActStatus
VAR_INPUT
    nAction : UINT;
END_VAR
CASE nAction OF
    GVL_Catalog.Cylinder_MoveTravail, GVL_Catalog.Cylinder_MoveRepos:
        _fMove := 0;
        _fSettle := 0;
        _nReached := 0;
        _OnStart := E_ActStatus.Busy;   // la commande est posée dans _OnCycle (attente si override 0 %)
    GVL_Catalog.Cylinder_LirePosition:
        _SetResult(1, _PositionCode());
        _OnStart := E_ActStatus.Done;
ELSE
    _OnStart := E_ActStatus.Error;
END_CASE
END_METHOD

METHOD PROTECTED _OnCycle : E_ActStatus
VAR_INPUT
    nAction : UINT;
END_VAR
VAR
    bTarget : BOOL;
    bSensorOk : BOOL;
    fCycleMs : LREAL;
END_VAR
fCycleMs := F_CycleMs();
IF _fEffOverride <= 0 AND _fMove = 0 THEN _OnCycle := E_ActStatus.Busy; RETURN; END_IF   // 0 % : on attend
bTarget := nAction = GVL_Catalog.Cylinder_MoveTravail;
_bCmdWork := bTarget;
_fMove := _fMove + fCycleMs;
// Capteur de départ toujours actif après 500 ms : vérin bloqué (erreur 102)
IF _fMove >= 500.0 AND ((bTarget AND _bHasRestSensor AND _bAtRest) OR (NOT bTarget AND _bHasWorkSensor AND _bAtWork)) THEN
    _Fail(GVL_Catalog.Cylinder_Err102, 0);
    _OnCycle := E_ActStatus.Error;
    RETURN;
END_IF
IF bTarget THEN
    bSensorOk := SEL(_bHasWorkSensor, _fMove >= _tNoSensorMs, _bAtWork AND NOT _bAtRest);
ELSE
    bSensorOk := SEL(_bHasRestSensor, _fMove >= _tNoSensorMs, _bAtRest AND NOT _bAtWork);
END_IF
IF bSensorOk THEN _fSettle := _fSettle + fCycleMs; ELSE _fSettle := 0; END_IF
IF _fSettle >= _tSettleMs THEN
    _nReached := SEL(bTarget, 1, 2);
    _OnCycle := E_ActStatus.Done;
ELSE
    _OnCycle := E_ActStatus.Busy;
END_IF
END_METHOD

METHOD PROTECTED _SafeState
CASE _eSafe OF
    0: _bCmdWork := FALSE;
    1: _bCmdWork := TRUE;
END_CASE                            // 2 : maintien
END_METHOD

METHOD PROTECTED _Monitor
IF _bAtWork AND _bAtRest THEN
    IF _eState <> E_ObjState.Error THEN _Fail(GVL_Catalog.Cylinder_Err100, 0); END_IF
ELSIF _eState = E_ObjState.Ready THEN
    // Perte du capteur de la position atteinte hors mouvement (erreur 101)
    IF (_nReached = 2 AND _bHasWorkSensor AND NOT _bAtWork) OR (_nReached = 1 AND _bHasRestSensor AND NOT _bAtRest) THEN
        _Fail(GVL_Catalog.Cylinder_Err101, _nReached);
        _nReached := 0;
    END_IF
END_IF
END_METHOD

METHOD PROTECTED _ReadHw
_bAtWork := F_ReadDI(_refCfg.aSignal[3]);
_bAtRest := F_ReadDI(_refCfg.aSignal[4]);
END_METHOD

METHOD PROTECTED _WriteHw
F_WriteDO(_refCfg.aSignal[1], _bCmdWork);
IF _bBistable THEN F_WriteDO(_refCfg.aSignal[2], NOT _bCmdWork); END_IF
END_METHOD

METHOD PROTECTED _Simulate
VAR
    fStep : LREAL;
END_VAR
fStep := F_CycleMs() / SEL(_refCfg.aParam[3] > 0, 300.0, _tNoSensorMs);
IF _bCmdWork THEN _fSimPos := MIN(1.0, _fSimPos + fStep); ELSE _fSimPos := MAX(0.0, _fSimPos - fStep); END_IF
_bAtWork := _fSimPos >= 1.0;
_bAtRest := _fSimPos <= 0.0;
IF _Forced(3) THEN _bAtWork := _ForcedValue(3) >= 0.5; END_IF
IF _Forced(4) THEN _bAtRest := _ForcedValue(4) >= 0.5; END_IF
END_METHOD

METHOD PRIVATE _PositionCode : LREAL
// 0 Inconnue, 1 Repos, 2 Travail, 3 Intermédiaire, 4 Incohérente
IF _bAtWork AND _bAtRest THEN
    _PositionCode := 4;
ELSIF _bAtRest THEN
    _PositionCode := 1;
ELSIF _bAtWork THEN
    _PositionCode := 2;
ELSIF _bHasWorkSensor OR _bHasRestSensor THEN
    _PositionCode := 3;
ELSE
    _PositionCode := 0;
END_IF
END_METHOD

METHOD PROTECTED _Publish
_stStatus.aValue[1] := _PositionCode();
IF _eState = E_ObjState.Busy THEN
    _stStatus.fProgress := LREAL_TO_REAL(MIN(1.0, _fMove / MAX(_tNoSensorMs, 1.0)));
END_IF
END_METHOD
END_FUNCTION_BLOCK

(* ---- FB_DigitalInput.st ---- *)
// Entrée numérique, type 1 (docs/03 § 3.1)
FUNCTION_BLOCK FB_DigitalInput EXTENDS FB_ObjectBase
VAR
    _bRaw : BOOL;                   // valeur lue (inversion P1 appliquée)
    _bValue : BOOL;                 // valeur filtrée (P2)
    _fDebounceMs : LREAL;
    _fChangeMs : LREAL;             // durée depuis laquelle la valeur lue diffère de la valeur filtrée
    _fWaitMs : LREAL;
END_VAR

METHOD PROTECTED _OnConfigure : BOOL
_fDebounceMs := LIMIT(0.0, _refCfg.aParam[2], 1000.0);
_OnConfigure := F_SignalValid(_refCfg.aSignal[1], E_SignalKind.DI);
END_METHOD

METHOD PROTECTED _OnStart : E_ActStatus
VAR_INPUT
    nAction : UINT;
END_VAR
_fWaitMs := 0;
CASE nAction OF
    GVL_Catalog.DigitalInput_Lire:
        _SetResult(1, BOOL_TO_LREAL(_bValue));
        _OnStart := E_ActStatus.Done;
    GVL_Catalog.DigitalInput_AttendreActif, GVL_Catalog.DigitalInput_AttendreInactif:
        _OnStart := _OnCycle(nAction);
ELSE
    _OnStart := E_ActStatus.Error;
END_CASE
END_METHOD

METHOD PROTECTED _OnCycle : E_ActStatus
VAR_INPUT
    nAction : UINT;
END_VAR
_fWaitMs := _fWaitMs + F_CycleMs();
// En simulation, sans forçage, l'attente se termine après 300 ms (docs/03 § 3.1)
IF _IsSimulated() AND NOT _Forced(1) AND _fWaitMs >= 300.0 THEN
    _bValue := nAction = GVL_Catalog.DigitalInput_AttendreActif;
END_IF
IF (nAction = GVL_Catalog.DigitalInput_AttendreActif) = _bValue THEN
    _OnCycle := E_ActStatus.Done;
ELSE
    _OnCycle := E_ActStatus.Busy;
END_IF
END_METHOD

METHOD PROTECTED _ReadHw
_bRaw := F_ReadDI(_refCfg.aSignal[1]) XOR (_refCfg.aParam[1] = 1);
_Debounce();
END_METHOD

METHOD PROTECTED _Simulate
IF _Forced(1) THEN
    _bRaw := _ForcedValue(1) >= 0.5;
    _Debounce();
END_IF
END_METHOD

METHOD PRIVATE _Debounce
IF _bRaw = _bValue THEN
    _fChangeMs := 0;
ELSE
    _fChangeMs := _fChangeMs + F_CycleMs();
    IF _fChangeMs >= _fDebounceMs THEN
        _bValue := _bRaw;
        _fChangeMs := 0;
    END_IF
END_IF
END_METHOD

METHOD PROTECTED _Publish
_stStatus.aValue[1] := BOOL_TO_LREAL(_bValue);
END_METHOD

PROPERTY Value : BOOL
GET
Value := _bValue;
END_GET
END_PROPERTY
END_FUNCTION_BLOCK

(* ---- FB_DigitalOutput.st ---- *)
// Sortie numérique, type 2 (docs/03 § 3.2)
FUNCTION_BLOCK FB_DigitalOutput EXTENDS FB_ObjectBase
VAR
    _bCmd : BOOL;
    _fPulseMs : LREAL;
    _fElapsed : LREAL;
END_VAR

METHOD PROTECTED _OnConfigure : BOOL
_OnConfigure := F_SignalValid(_refCfg.aSignal[1], E_SignalKind.DO);
END_METHOD

METHOD PROTECTED _DefaultTimeoutMs : UDINT
VAR_INPUT
    nAction : UINT;
END_VAR
IF nAction = GVL_Catalog.DigitalOutput_Impulsion THEN
    _DefaultTimeoutMs := LREAL_TO_UDINT(_ParamReal(1, _refCfg.aParam[2])) + 1000;
ELSE
    _DefaultTimeoutMs := 0;
END_IF
END_METHOD

METHOD PROTECTED _ValidateParams : BOOL
VAR_INPUT
    nAction : UINT;
END_VAR
_ValidateParams := nAction <> GVL_Catalog.DigitalOutput_Impulsion OR _ParamReal(1, _refCfg.aParam[2]) >= 1.0;
END_METHOD

METHOD PROTECTED _OnStart : E_ActStatus
VAR_INPUT
    nAction : UINT;
END_VAR
CASE nAction OF
    GVL_Catalog.DigitalOutput_Activer:
        _bCmd := TRUE;
        _OnStart := E_ActStatus.Done;
    GVL_Catalog.DigitalOutput_Desactiver:
        _bCmd := FALSE;
        _OnStart := E_ActStatus.Done;
    GVL_Catalog.DigitalOutput_Impulsion:
        _fPulseMs := LIMIT(1.0, _ParamReal(1, _refCfg.aParam[2]), 60000.0);
        _fElapsed := 0;
        _bCmd := TRUE;
        _OnStart := E_ActStatus.Busy;
ELSE
    _OnStart := E_ActStatus.Error;
END_CASE
END_METHOD

METHOD PROTECTED _OnCycle : E_ActStatus
VAR_INPUT
    nAction : UINT;
END_VAR
_fElapsed := _fElapsed + F_CycleMs();
IF _fElapsed >= _fPulseMs THEN
    _bCmd := FALSE;
    _OnCycle := E_ActStatus.Done;
ELSE
    _OnCycle := E_ActStatus.Busy;
END_IF
END_METHOD

METHOD PROTECTED _SafeState
CASE LREAL_TO_INT(_refCfg.aParam[3]) OF
    0: _bCmd := FALSE;
    1: _bCmd := TRUE;
END_CASE                            // 2 : maintien
END_METHOD

METHOD PROTECTED _WriteHw
F_WriteDO(_refCfg.aSignal[1], _bCmd XOR (_refCfg.aParam[1] = 1));
END_METHOD

METHOD PROTECTED _Publish
_stStatus.aValue[1] := BOOL_TO_LREAL(_bCmd);
END_METHOD
END_FUNCTION_BLOCK

(* ---- FB_Gripper.st ---- *)
// Pince, type 21 (docs/03 § 5.2). Seul le pneumatique est réalisé ; l'électrique (P1 = 2) attend son interface :
// la configuration est alors refusée.
FUNCTION_BLOCK FB_Gripper EXTENDS FB_ObjectBase
VAR
    _bBistable : BOOL;
    _bCmdClose : BOOL;
    _bClosed : BOOL;
    _bOpen : BOOL;
    _bPart : BOOL;
    _bHasClosed : BOOL;
    _bHasOpen : BOOL;
    _bHasPart : BOOL;
    _bHolding : BOOL;               // fermée sur pièce : une perte de pièce est une erreur 101
    _fMove : LREAL;
    _fSimPos : LREAL;               // 0 ouverte, 1 fermée
    _bSimPart : BOOL := TRUE;       // simulation : une pièce est présente entre les doigts
END_VAR

METHOD PROTECTED _OnConfigure : BOOL
_bBistable := _refCfg.aParam[1] = 1;
_bHasClosed := F_SignalValid(_refCfg.aSignal[3], E_SignalKind.DI);
_bHasOpen := F_SignalValid(_refCfg.aSignal[4], E_SignalKind.DI);
_bHasPart := F_SignalValid(_refCfg.aSignal[5], E_SignalKind.DI);
_bHolding := FALSE;
_OnConfigure := _refCfg.aParam[1] < 2
                AND F_SignalValid(_refCfg.aSignal[1], E_SignalKind.DO)
                AND (NOT _bBistable OR F_SignalValid(_refCfg.aSignal[2], E_SignalKind.DO));
END_METHOD

METHOD PROTECTED _OnStart : E_ActStatus
VAR_INPUT
    nAction : UINT;
END_VAR
_fMove := 0;
CASE nAction OF
    GVL_Catalog.Gripper_Ouvrir:
        _bCmdClose := FALSE;
        _bHolding := FALSE;
        _OnStart := E_ActStatus.Busy;
    GVL_Catalog.Gripper_Fermer, GVL_Catalog.Gripper_SerrerSurPiece:
        _bCmdClose := TRUE;
        _OnStart := E_ActStatus.Busy;
    GVL_Catalog.Gripper_VerifierPresencePiece:
        _SetResult(1, BOOL_TO_LREAL(_PartPresent()));
        _OnStart := E_ActStatus.Done;
ELSE
    _OnStart := E_ActStatus.Error;
END_CASE
END_METHOD

METHOD PROTECTED _OnCycle : E_ActStatus
VAR_INPUT
    nAction : UINT;
END_VAR
VAR
    bReached : BOOL;
END_VAR
_fMove := _fMove + F_CycleMs();
IF _bCmdClose THEN
    bReached := SEL(_bHasClosed, _fMove >= _refCfg.aParam[2], _bClosed);
ELSE
    bReached := SEL(_bHasOpen, _fMove >= _refCfg.aParam[2], _bOpen);
END_IF
IF NOT bReached THEN
    _OnCycle := E_ActStatus.Busy;
    RETURN;
END_IF
IF nAction = GVL_Catalog.Gripper_SerrerSurPiece THEN
    _SetResult(1, BOOL_TO_LREAL(_PartPresent()));
    IF NOT _PartPresent() THEN
        _Fail(GVL_Catalog.Gripper_Err100, 0);       // pièce absente à la fermeture
        _OnCycle := E_ActStatus.Error;
        RETURN;
    END_IF
    _bHolding := TRUE;
END_IF
_OnCycle := E_ActStatus.Done;
END_METHOD

METHOD PRIVATE _PartPresent : BOOL
// Avec un capteur de présence : le capteur ; sinon, fermée sans atteindre la butée « fermée » = sur pièce
IF _bHasPart THEN
    _PartPresent := _bPart;
ELSE
    _PartPresent := _bCmdClose AND NOT _bOpen;
END_IF
END_METHOD

METHOD PROTECTED _Monitor
IF _bHasClosed AND _bHasOpen AND _bClosed AND _bOpen THEN
    IF _eState <> E_ObjState.Error THEN _Fail(GVL_Catalog.Gripper_Err102, 0); END_IF
ELSIF _bHolding AND _bHasPart AND NOT _bPart AND _eState <> E_ObjState.Error THEN
    _bHolding := FALSE;
    _Fail(GVL_Catalog.Gripper_Err101, 0);          // pièce perdue pendant le maintien
END_IF
END_METHOD

// État sûr : maintien (docs/03, catalogue)
METHOD PROTECTED _SafeState
;
END_METHOD

METHOD PROTECTED _ReadHw
_bClosed := F_ReadDI(_refCfg.aSignal[3]);
_bOpen := F_ReadDI(_refCfg.aSignal[4]);
_bPart := F_ReadDI(_refCfg.aSignal[5]);
END_METHOD

METHOD PROTECTED _Simulate
VAR
    fStep : LREAL;
END_VAR
fStep := F_CycleMs() / MAX(_refCfg.aParam[2], 10.0);
IF _bCmdClose THEN _fSimPos := MIN(1.0, _fSimPos + fStep); ELSE _fSimPos := MAX(0.0, _fSimPos - fStep); END_IF
_bOpen := _fSimPos <= 0.0;
_bClosed := _fSimPos >= 1.0;
_bPart := _bSimPart AND _bCmdClose AND _fSimPos >= 1.0;
IF _Forced(3) THEN _bClosed := _ForcedValue(3) >= 0.5; END_IF
IF _Forced(4) THEN _bOpen := _ForcedValue(4) >= 0.5; END_IF
IF _Forced(5) THEN _bPart := _ForcedValue(5) >= 0.5; END_IF
END_METHOD

METHOD PROTECTED _WriteHw
F_WriteDO(_refCfg.aSignal[1], _bCmdClose);
IF _bBistable THEN F_WriteDO(_refCfg.aSignal[2], NOT _bCmdClose); END_IF
END_METHOD

METHOD PROTECTED _Publish
// 0 Inconnu, 1 Ouverte, 2 Fermée, 3 Fermée sur pièce
IF _bCmdClose AND _PartPresent() THEN
    _stStatus.aValue[1] := 3;
ELSIF _bCmdClose AND (_bClosed OR NOT _bHasClosed) THEN
    _stStatus.aValue[1] := 2;
ELSIF NOT _bCmdClose AND (_bOpen OR NOT _bHasOpen) THEN
    _stStatus.aValue[1] := 1;
ELSE
    _stStatus.aValue[1] := 0;
END_IF
_stStatus.aValue[2] := BOOL_TO_LREAL(_PartPresent());
END_METHOD
END_FUNCTION_BLOCK

(* ---- FB_Group.st ---- *)
// Module libre et base des modules, type 100 (docs/03 § 9.1) : override commun et état agrégé de ses enfants
FUNCTION_BLOCK FB_Group EXTENDS FB_ObjectBase IMPLEMENTS I_Group
VAR
    _eAggregate : E_ObjState := E_ObjState.Ready;
END_VAR

METHOD SetAggregate
VAR_INPUT
    eState : E_ObjState;
END_VAR
_eAggregate := eState;
END_METHOD

PROPERTY NodeState : E_ObjState
GET
IF _eState = E_ObjState.Disabled THEN
    NodeState := E_ObjState.Disabled;
ELSE
    NodeState := _eAggregate;
END_IF
END_GET
END_PROPERTY

METHOD PROTECTED _OnStart : E_ActStatus
VAR_INPUT
    nAction : UINT;
END_VAR
_OnStart := E_ActStatus.Error;      // un module n'a pas d'action : ses fonctions sont dépliées par le compilateur
END_METHOD
END_FUNCTION_BLOCK

(* ---- FB_KeyenceGT2.st ---- *)
// Palpeur Keyence GT2, type 31 (docs/03 § 6.2), mode signaux : S1 AI valeur. Le mode réseau (P1 = 1) n'est pas
// encore écrit : la configuration est refusée.
// Hypothèse : la valeur brute de l'entrée analogique est en micromètres (1 = 0,001 mm), comme la sortie
// analogique du GT2 réglée sur ±32 mm. À confirmer avec le câblage réel.
FUNCTION_BLOCK FB_KeyenceGT2 EXTENDS FB_ObjectBase
VAR
    _fValue : LREAL;                // mm, après remise à zéro
    _fRaw : LREAL;                  // mm, avant remise à zéro
    _fZero : LREAL;
    _bOutOfRange : BOOL;
    _fStabMs : LREAL;
    _nWanted : INT;
    _nTaken : INT;
    _fSum : LREAL;
    _fSimValue : LREAL;
END_VAR
VAR PERSISTENT
    _fZeroKept : LREAL;             // remise à zéro gardée après une coupure
END_VAR

METHOD PROTECTED _OnConfigure : BOOL
IF _bNewObject THEN _fZeroKept := 0; END_IF
_fZero := _fZeroKept;
_fSimValue := _refCfg.aParam[2];
_OnConfigure := _refCfg.aParam[1] = 0 AND F_SignalValid(_refCfg.aSignal[1], E_SignalKind.AI);
END_METHOD

METHOD PROTECTED _OnStart : E_ActStatus
VAR_INPUT
    nAction : UINT;
END_VAR
CASE nAction OF
    GVL_Catalog.KeyenceGT2_Mesurer:
        _nWanted := LIMIT(1, LREAL_TO_INT(_ParamReal(1, _refCfg.aParam[5])), 1000);
        _nTaken := 0;
        _fSum := 0;
        _fStabMs := 0;
        _OnStart := E_ActStatus.Busy;
    GVL_Catalog.KeyenceGT2_RemiseAZero:
        _fZero := _fRaw;
        _fZeroKept := _fZero;
        _OnStart := E_ActStatus.Done;
    GVL_Catalog.KeyenceGT2_LireValeurCourante:
        _SetResult(1, _fValue);
        _OnStart := E_ActStatus.Done;
ELSE
    _OnStart := E_ActStatus.Error;
END_CASE
END_METHOD

METHOD PROTECTED _OnCycle : E_ActStatus
VAR_INPUT
    nAction : UINT;
END_VAR
VAR
    fMean : LREAL;
    fHigh : LREAL;
    fLow : LREAL;
END_VAR
_OnCycle := E_ActStatus.Busy;
IF _bOutOfRange THEN
    _Fail(GVL_Catalog.KeyenceGT2_Err100, 0);
    _OnCycle := E_ActStatus.Error;
    RETURN;
END_IF
// Stabilisation P6, puis un échantillon par cycle
_fStabMs := _fStabMs + F_CycleMs();
IF _fStabMs < MAX(0.0, _refCfg.aParam[6]) THEN RETURN; END_IF
_fSum := _fSum + _fValue;
_nTaken := _nTaken + 1;
IF _nTaken < _nWanted THEN RETURN; END_IF
fMean := _fSum / INT_TO_LREAL(_nTaken);
fHigh := _refCfg.aParam[2] + ABS(_refCfg.aParam[3]);
fLow := _refCfg.aParam[2] - ABS(_refCfg.aParam[4]);
_SetResult(1, fMean);
IF fMean > fHigh THEN
    _SetJudgement(2, E_Judgement.High);
ELSIF fMean < fLow THEN
    _SetJudgement(2, E_Judgement.Low);
ELSE
    _SetJudgement(2, E_Judgement.Ok);
END_IF
_OnCycle := E_ActStatus.Done;
END_METHOD

METHOD PROTECTED _ReadHw
VAR
    nRaw : INT;
END_VAR
nRaw := F_ReadAI(_refCfg.aSignal[1]);
_bOutOfRange := nRaw = 32767 OR nRaw = -32768;
_fRaw := INT_TO_LREAL(nRaw) * 0.001;
_fValue := _fRaw - _fZero;
END_METHOD

// Simulation : valeur de référence P2 avec un bruit de ±10 % de la tolérance haute (docs/03 § 6.2)
METHOD PROTECTED _Simulate
_fRaw := _fSimValue + (F_SimRandom() - 0.5) * 0.2 * ABS(_refCfg.aParam[3]) + _fZero;
IF _Forced(1) THEN _fRaw := _ForcedValue(1) + _fZero; END_IF       // valeur forcée en mm
_bOutOfRange := FALSE;
_fValue := _fRaw - _fZero;
END_METHOD

METHOD PROTECTED _Publish
_stStatus.aValue[1] := _fValue;
END_METHOD
END_FUNCTION_BLOCK

(* ---- FB_KeyenceIV.st ---- *)
// Vision Keyence IV, type 30 (docs/03 § 6.1), mode signaux : S1 DO déclenchement, S2 DI prêt, S3 DI résultat OK,
// S4 DI résultat NOK. Le mode réseau (P1 = 1) n'est pas encore écrit : la configuration est refusée.
// Hypothèse : en mode signaux, le programme ne se change pas par les signaux ; « Sélectionner programme »
// mémorise le n° demandé (affiché, rendu par la HMI) sans le transmettre à l'appareil.
FUNCTION_BLOCK FB_KeyenceIV EXTENDS FB_ObjectBase
VAR
    _bTrigger : BOOL;
    _bReady : BOOL;
    _bOk : BOOL;
    _bNok : BOOL;
    _fWaitMs : LREAL;
    _nProgram : INT;
    _eLast : E_Judgement;
    _fLastValue : LREAL;
    _bSimResult : BOOL;             // simulation : un résultat est présent
    _bSimOk : BOOL;
END_VAR

METHOD PROTECTED _OnConfigure : BOOL
_nProgram := LREAL_TO_INT(_refCfg.aParam[2]);
_OnConfigure := _refCfg.aParam[1] = 0
                AND F_SignalValid(_refCfg.aSignal[1], E_SignalKind.DO)
                AND F_SignalValid(_refCfg.aSignal[3], E_SignalKind.DI)
                AND F_SignalValid(_refCfg.aSignal[4], E_SignalKind.DI);
END_METHOD

METHOD PROTECTED _OnStart : E_ActStatus
VAR_INPUT
    nAction : UINT;
END_VAR
CASE nAction OF
    GVL_Catalog.KeyenceIV_SelectionnerProgramme:
        _nProgram := LREAL_TO_INT(_ParamReal(1, _refCfg.aParam[2]));
        _OnStart := E_ActStatus.Done;
    GVL_Catalog.KeyenceIV_Declencher:
        IF F_SignalValid(_refCfg.aSignal[2], E_SignalKind.DI) AND NOT _bReady THEN
            _Fail(GVL_Catalog.KeyenceIV_Err100, 0);
            _OnStart := E_ActStatus.Error;
            RETURN;
        END_IF
        _fWaitMs := 0;
        _bTrigger := TRUE;
        _bSimResult := FALSE;
        _OnStart := E_ActStatus.Busy;
    GVL_Catalog.KeyenceIV_LireDernierResultat:
        _SetJudgement(1, _eLast);
        _SetResult(2, _fLastValue);
        _OnStart := E_ActStatus.Done;
ELSE
    _OnStart := E_ActStatus.Error;
END_CASE
END_METHOD

METHOD PROTECTED _OnCycle : E_ActStatus
VAR_INPUT
    nAction : UINT;
END_VAR
_OnCycle := E_ActStatus.Busy;
_fWaitMs := _fWaitMs + F_CycleMs();
// Le résultat est lu après l'attente P3, quand l'une des deux sorties du capteur est active
IF _fWaitMs < MAX(0.0, _refCfg.aParam[3]) OR NOT (_bOk XOR _bNok) THEN RETURN; END_IF
_bTrigger := FALSE;
IF _bOk THEN _eLast := E_Judgement.Ok; ELSE _eLast := E_Judgement.Nok; END_IF
_fLastValue := 0;                   // pas de valeur mesurée en mode signaux
_SetJudgement(1, _eLast);
_SetResult(2, _fLastValue);
_OnCycle := E_ActStatus.Done;
END_METHOD

METHOD PROTECTED _OnAbort
VAR_INPUT
    nAction : UINT;
END_VAR
_bTrigger := FALSE;
END_METHOD

METHOD PROTECTED _SafeState
_bTrigger := FALSE;
END_METHOD

METHOD PROTECTED _ReadHw
_bReady := F_ReadDI(_refCfg.aSignal[2]);
_bOk := F_ReadDI(_refCfg.aSignal[3]);
_bNok := F_ReadDI(_refCfg.aSignal[4]);
END_METHOD

METHOD PROTECTED _WriteHw
F_WriteDO(_refCfg.aSignal[1], _bTrigger);
END_METHOD

// Simulation : prêt ; à chaque déclenchement, jugement bon avec une probabilité de 95 % (docs/03 § 6.1)
METHOD PROTECTED _Simulate
IF _bTrigger AND NOT _bSimResult THEN
    _bSimResult := TRUE;
    _bSimOk := F_SimRandom() < 0.95;
END_IF
_bReady := TRUE;
_bOk := _bSimResult AND _bSimOk;
_bNok := _bSimResult AND NOT _bSimOk;
IF _Forced(2) THEN _bReady := _ForcedValue(2) >= 0.5; END_IF
IF _Forced(3) THEN _bOk := _ForcedValue(3) >= 0.5; END_IF
IF _Forced(4) THEN _bNok := _ForcedValue(4) >= 0.5; END_IF
END_METHOD

METHOD PROTECTED _Publish
_stStatus.aValue[1] := TO_LREAL(_eLast);
_stStatus.aValue[2] := INT_TO_LREAL(_nProgram);
END_METHOD
END_FUNCTION_BLOCK

(* ---- FB_Light.st ---- *)
// Éclairage, type 35 (docs/03 § 6.6) : S1 DO commande, S2 AO intensité (optionnel, 0 à 100 % = 0 à 32767),
// S3 DO synchronisation caméra (optionnel, active pendant un flash). État sûr : éteint.
FUNCTION_BLOCK FB_Light EXTENDS FB_ObjectBase
VAR
    _bOn : BOOL;
    _bSync : BOOL;
    _fIntensity : LREAL;            // %
    _fFlashMs : LREAL;
    _fElapsed : LREAL;
END_VAR

METHOD PROTECTED _OnConfigure : BOOL
_fIntensity := LIMIT(0.0, _refCfg.aParam[2], 100.0);
_OnConfigure := F_SignalValid(_refCfg.aSignal[1], E_SignalKind.DO);
END_METHOD

METHOD PROTECTED _DefaultTimeoutMs : UDINT
VAR_INPUT
    nAction : UINT;
END_VAR
IF nAction = GVL_Catalog.Light_Flasher THEN
    _DefaultTimeoutMs := LREAL_TO_UDINT(MAX(0.0, _ParamReal(1, _refCfg.aParam[3]))) + 200;
ELSE
    _DefaultTimeoutMs := 0;
END_IF
END_METHOD

METHOD PROTECTED _OnStart : E_ActStatus
VAR_INPUT
    nAction : UINT;
END_VAR
CASE nAction OF
    GVL_Catalog.Light_Allumer:
        _fIntensity := LIMIT(0.0, _ParamReal(1, _refCfg.aParam[2]), 100.0);
        _bOn := TRUE;
        _OnStart := E_ActStatus.Done;
    GVL_Catalog.Light_Eteindre:
        _bOn := FALSE;
        _bSync := FALSE;
        _OnStart := E_ActStatus.Done;
    GVL_Catalog.Light_ReglerIntensite:
        _fIntensity := LIMIT(0.0, _ParamReal(1, _fIntensity), 100.0);
        _OnStart := E_ActStatus.Done;
    GVL_Catalog.Light_Flasher:
        _fFlashMs := MAX(0.0, _ParamReal(1, _refCfg.aParam[3]));
        _fIntensity := LIMIT(0.0, _ParamReal(2, _refCfg.aParam[2]), 100.0);
        _fElapsed := 0;
        _bOn := TRUE;
        _bSync := TRUE;
        _OnStart := E_ActStatus.Busy;
ELSE
    _OnStart := E_ActStatus.Error;
END_CASE
END_METHOD

METHOD PROTECTED _OnCycle : E_ActStatus
VAR_INPUT
    nAction : UINT;
END_VAR
_fElapsed := _fElapsed + F_CycleMs();
IF _fElapsed >= _fFlashMs THEN
    _bOn := FALSE;
    _bSync := FALSE;
    _OnCycle := E_ActStatus.Done;
ELSE
    _OnCycle := E_ActStatus.Busy;
END_IF
END_METHOD

METHOD PROTECTED _OnAbort
VAR_INPUT
    nAction : UINT;
END_VAR
_bOn := FALSE;
_bSync := FALSE;
END_METHOD

METHOD PROTECTED _SafeState
_bOn := FALSE;
_bSync := FALSE;
END_METHOD

METHOD PROTECTED _WriteHw
F_WriteDO(_refCfg.aSignal[1], _bOn);
F_WriteAO(_refCfg.aSignal[2], LREAL_TO_INT(_fIntensity * 32767.0 / 100.0));
F_WriteDO(_refCfg.aSignal[3], _bSync);
END_METHOD

METHOD PROTECTED _Publish
_stStatus.aValue[1] := SEL(_bOn, 0.0, 1.0);
_stStatus.aValue[2] := _fIntensity;
END_METHOD
END_FUNCTION_BLOCK

(* ---- FB_Magazine.st ---- *)
// Palettiseur ou magasin, type 45 (docs/03 § 7.6) : S1 DI plateau présent, S2 DI magasin vide, S3 DI magasin
// plein, S4 DO présenter, S5 DO évacuer. Cases numérotées ligne par ligne depuis la première case (position
// nommée P5 de la station), pas P3 en X et P4 en Y. L'occupation du plateau présent est persistante.
FUNCTION_BLOCK FB_Magazine EXTENDS FB_ObjectBase
VAR
    _bPresent : BOOL;
    _bEmpty : BOOL;
    _bFull : BOOL;
    _bCmdPresent : BOOL;
    _bCmdEvacuate : BOOL;
    _nRows : INT;
    _nCols : INT;
    _fSimMs : LREAL;
    _bSimPresent : BOOL;
END_VAR
VAR PERSISTENT
    _aOccupied : ARRAY[1..256] OF BOOL;
END_VAR

METHOD PROTECTED _OnConfigure : BOOL
_nRows := LIMIT(1, LREAL_TO_INT(_refCfg.aParam[1]), 16);
_nCols := LIMIT(1, LREAL_TO_INT(_refCfg.aParam[2]), 16);
IF _bNewObject THEN MEMSET(ADR(_aOccupied), 0, SIZEOF(_aOccupied)); END_IF
_OnConfigure := F_SignalValid(_refCfg.aSignal[1], E_SignalKind.DI)
                AND F_SignalValid(_refCfg.aSignal[4], E_SignalKind.DO)
                AND F_SignalValid(_refCfg.aSignal[5], E_SignalKind.DO);
END_METHOD

METHOD PROTECTED _OnStart : E_ActStatus
VAR_INPUT
    nAction : UINT;
END_VAR
VAR
    n : INT;
END_VAR
CASE nAction OF
    GVL_Catalog.Magazine_PresenterPlateauSuivant:
        IF _bEmpty THEN _Fail(GVL_Catalog.Magazine_Err100, 0); _OnStart := E_ActStatus.Error; RETURN; END_IF
        _bCmdPresent := TRUE;
        _fSimMs := 0;
        _OnStart := E_ActStatus.Busy;
    GVL_Catalog.Magazine_EvacuerPlateau:
        IF NOT _bPresent THEN _Fail(GVL_Catalog.Magazine_Err102, 0); _OnStart := E_ActStatus.Error; RETURN; END_IF
        IF _bFull THEN _Fail(GVL_Catalog.Magazine_Err101, 0); _OnStart := E_ActStatus.Error; RETURN; END_IF
        _bCmdEvacuate := TRUE;
        _fSimMs := 0;
        _OnStart := E_ActStatus.Busy;
    GVL_Catalog.Magazine_PositionDeLaCase:
        n := LREAL_TO_INT(_ParamReal(1, 0));
        IF n = 0 THEN n := _FirstFree(); END_IF
        IF n < 1 OR n > _nRows * _nCols THEN _Fail(GVL_Catalog.Err_BadParam, 1); _OnStart := E_ActStatus.Error; RETURN; END_IF
        _SetResultPos(1, _CellPos(n));
        _SetResult(2, INT_TO_LREAL(n));
        _OnStart := E_ActStatus.Done;
    GVL_Catalog.Magazine_MarquerCase:
        n := LREAL_TO_INT(_ParamReal(1, 0));
        IF n < 1 OR n > _nRows * _nCols THEN _Fail(GVL_Catalog.Err_BadParam, 1); _OnStart := E_ActStatus.Error; RETURN; END_IF
        _aOccupied[n] := _ParamReal(2, 1) <> 0;
        _OnStart := E_ActStatus.Done;
    GVL_Catalog.Magazine_LireOccupation:
        n := _CountOccupied();
        _SetResult(1, INT_TO_LREAL(n));
        _SetResult(2, INT_TO_LREAL(_nRows * _nCols - n));
        _SetResult(3, SEL(n >= _nRows * _nCols, 0.0, 1.0));
        _OnStart := E_ActStatus.Done;
ELSE
    _OnStart := E_ActStatus.Error;
END_CASE
END_METHOD

METHOD PROTECTED _OnCycle : E_ActStatus
VAR_INPUT
    nAction : UINT;
END_VAR
_OnCycle := E_ActStatus.Busy;
CASE nAction OF
    GVL_Catalog.Magazine_PresenterPlateauSuivant:
        IF _bPresent THEN
            _bCmdPresent := FALSE;
            MEMSET(ADR(_aOccupied), 0, SIZEOF(_aOccupied));        // plateau neuf : toutes les cases libres
            _OnCycle := E_ActStatus.Done;
        ELSIF _fElapsedMs + 100.0 >= UDINT_TO_LREAL(_nTimeoutMs) AND _nTimeoutMs > 0 THEN
            _bCmdPresent := FALSE;
            _Fail(GVL_Catalog.Magazine_Err102, 0);
            _OnCycle := E_ActStatus.Error;
        END_IF
    GVL_Catalog.Magazine_EvacuerPlateau:
        IF NOT _bPresent THEN
            _bCmdEvacuate := FALSE;
            _OnCycle := E_ActStatus.Done;
        ELSIF _fElapsedMs + 100.0 >= UDINT_TO_LREAL(_nTimeoutMs) AND _nTimeoutMs > 0 THEN
            _bCmdEvacuate := FALSE;
            _Fail(GVL_Catalog.Magazine_Err103, 0);
            _OnCycle := E_ActStatus.Error;
        END_IF
ELSE
    _OnCycle := E_ActStatus.Done;
END_CASE
END_METHOD

METHOD PROTECTED _OnAbort
VAR_INPUT
    nAction : UINT;
END_VAR
_bCmdPresent := FALSE;
_bCmdEvacuate := FALSE;
END_METHOD

METHOD PROTECTED _SafeState
_bCmdPresent := FALSE;
_bCmdEvacuate := FALSE;
END_METHOD

METHOD PROTECTED _ReadHw
_bPresent := F_ReadDI(_refCfg.aSignal[1]);
_bEmpty := F_ReadDI(_refCfg.aSignal[2]);
_bFull := F_ReadDI(_refCfg.aSignal[3]);
END_METHOD

METHOD PROTECTED _WriteHw
F_WriteDO(_refCfg.aSignal[4], _bCmdPresent);
F_WriteDO(_refCfg.aSignal[5], _bCmdEvacuate);
END_METHOD

// Simulation : un plateau arrive ou part 1 s après la commande ; le magasin n'est jamais vide ni plein
METHOD PROTECTED _Simulate
IF _bCmdPresent OR _bCmdEvacuate THEN _fSimMs := _fSimMs + F_CycleMs(); END_IF
IF _bCmdPresent AND _fSimMs >= 1000.0 THEN _bSimPresent := TRUE; END_IF
IF _bCmdEvacuate AND _fSimMs >= 1000.0 THEN _bSimPresent := FALSE; END_IF
_bPresent := _bSimPresent;
_bEmpty := FALSE;
_bFull := FALSE;
IF _Forced(1) THEN _bPresent := _ForcedValue(1) >= 0.5; END_IF
IF _Forced(2) THEN _bEmpty := _ForcedValue(2) >= 0.5; END_IF
IF _Forced(3) THEN _bFull := _ForcedValue(3) >= 0.5; END_IF
END_METHOD

METHOD PRIVATE _FirstFree : INT
VAR
    i : INT;
END_VAR
_FirstFree := 0;
FOR i := 1 TO _nRows * _nCols DO
    IF NOT _aOccupied[i] THEN _FirstFree := i; RETURN; END_IF
END_FOR
END_METHOD

METHOD PRIVATE _CountOccupied : INT
VAR
    i : INT;
END_VAR
_CountOccupied := 0;
FOR i := 1 TO _nRows * _nCols DO
    IF _aOccupied[i] THEN _CountOccupied := _CountOccupied + 1; END_IF
END_FOR
END_METHOD

// Position de la case n : première case (position nommée P5 de la station) + décalage de colonne et de ligne
METHOD PRIVATE _CellPos : ST_Position
VAR_INPUT
    n : INT;
END_VAR
VAR
    nPos : INT;
END_VAR
nPos := LREAL_TO_INT(_refCfg.aParam[5]);
IF _stInfo.nStation >= 1 AND _stInfo.nStation <= GVL_Const.MAX_STATIONS AND nPos >= 1 AND nPos <= GVL_Const.MAX_NAMED_POS THEN
    _CellPos := GVL_Active.aStation[_stInfo.nStation].aPos[nPos].stPos;
END_IF
_CellPos.fX := _CellPos.fX + INT_TO_LREAL((n - 1) MOD _nCols) * _refCfg.aParam[3];
_CellPos.fY := _CellPos.fY + INT_TO_LREAL((n - 1) / _nCols) * _refCfg.aParam[4];
END_METHOD

METHOD PROTECTED _Publish
_stStatus.aValue[1] := SEL(_bPresent, 0.0, 1.0);
_stStatus.aValue[2] := INT_TO_LREAL(_CountOccupied());
END_METHOD
END_FUNCTION_BLOCK

(* ---- FB_PlanarMover.st ---- *)
// Mover, type 14, niveau machine (docs/03 § 4.4) : mode manuel des movers (docs/05 § 6.5). L'élément matériel
// D est le n° du mover ; les mouvements passent par le gestionnaire de movers (GVL_IoRef.ipMovers), qui tient
// l'occupation des positions planaires à jour.
FUNCTION_BLOCK FB_PlanarMover EXTENDS FB_ObjectBase
VAR
    _nMover : USINT;
    _stTarget : ST_Position;
    _stLast : ST_Position;
    _fSpeed : LREAL;                // mm/s, estimée d'un cycle à l'autre
END_VAR

METHOD PROTECTED _OnConfigure : BOOL
_nMover := INT_TO_USINT(LIMIT(0, _refCfg.nDevice, GVL_Const.MAX_MOVERS));
_OnConfigure := _nMover >= 1;
END_METHOD

METHOD PROTECTED _OnStart : E_ActStatus
VAR_INPUT
    nAction : UINT;
END_VAR
VAR
    fPct : LREAL := 100.0;
END_VAR
IF GVL_IoRef.ipMovers = 0 THEN
    _Fail(GVL_Catalog.Err_NotWired, 0);
    _OnStart := E_ActStatus.Error;
    RETURN;
END_IF
CASE nAction OF
    GVL_Catalog.PlanarMover_MoveVersPosition:
        IF _stParams.aKind[1] <> E_ParamKind.Position THEN
            _Fail(GVL_Catalog.Err_BadParam, 1);
            _OnStart := E_ActStatus.Error;
            RETURN;
        END_IF
        _stTarget := _stParams.stPos;
        IF _stParams.aKind[2] = E_ParamKind.SpeedPercent OR _stParams.aKind[2] = E_ParamKind.Real THEN fPct := _stParams.aReal[2]; END_IF
        IF NOT GVL_IoRef.ipMovers.MoveFree(_nMover, _stTarget, fPct * _fEffOverride / 100.0) THEN
            _Fail(GVL_Catalog.Err_NotReady, 0);         // position tenue par un autre mover, ou système inactif
            _OnStart := E_ActStatus.Error;
            RETURN;
        END_IF
        _OnStart := E_ActStatus.Busy;
    GVL_Catalog.PlanarMover_Stop:
        GVL_IoRef.ipMovers.StopMover(_nMover);
        _OnStart := E_ActStatus.Done;
    GVL_Catalog.PlanarMover_LirePosition:
        _SetResultPos(1, GVL_IoRef.ipMovers.Position(_nMover));
        _OnStart := E_ActStatus.Done;
ELSE
    _OnStart := E_ActStatus.Error;
END_CASE
END_METHOD

METHOD PROTECTED _OnCycle : E_ActStatus
VAR_INPUT
    nAction : UINT;
END_VAR
VAR
    stPos : ST_Position;
END_VAR
_OnCycle := E_ActStatus.Busy;
IF nAction <> GVL_Catalog.PlanarMover_MoveVersPosition THEN _OnCycle := E_ActStatus.Done; RETURN; END_IF
stPos := GVL_IoRef.ipMovers.Position(_nMover);
IF NOT GVL_IoRef.ipMovers.Moving(_nMover) THEN
    IF ABS(stPos.fX - _stTarget.fX) <= 0.5 AND ABS(stPos.fY - _stTarget.fY) <= 0.5 THEN
        _OnCycle := E_ActStatus.Done;
    ELSE
        _Fail(GVL_Catalog.Err_Aborted, 0);              // arrêté avant la cible (collision, arrêt du système)
        _OnCycle := E_ActStatus.Error;
    END_IF
END_IF
END_METHOD

METHOD PROTECTED _OnAbort
VAR_INPUT
    nAction : UINT;
END_VAR
IF GVL_IoRef.ipMovers <> 0 THEN GVL_IoRef.ipMovers.StopMover(_nMover); END_IF
END_METHOD

METHOD PROTECTED _Publish
VAR
    stPos : ST_Position;
    fDt : LREAL;
END_VAR
IF GVL_IoRef.ipMovers = 0 THEN RETURN; END_IF
stPos := GVL_IoRef.ipMovers.Position(_nMover);
fDt := F_CycleMs();
IF fDt > 0 THEN _fSpeed := SQRT(EXPT(stPos.fX - _stLast.fX, 2) + EXPT(stPos.fY - _stLast.fY, 2)) * 1000.0 / fDt; END_IF
_stLast := stPos;
_stStatus.aValue[1] := stPos.fX;
_stStatus.aValue[2] := stPos.fY;
_stStatus.aValue[3] := stPos.fC;
_stStatus.aValue[4] := _fSpeed;
END_METHOD
END_FUNCTION_BLOCK

(* ---- FB_PlanarSystem.st ---- *)
// Système planaire, type 13, niveau machine (docs/03 § 4.3) : activation, désactivation, acquittement du pilote
// planaire (GVL_IoRef.ipPlanar). Les erreurs du système (100 à 102) sont levées par FB_Machine, qui tient l'état.
FUNCTION_BLOCK FB_PlanarSystem EXTENDS FB_ObjectBase
VAR
    _nDetected : INT;
END_VAR

METHOD PROTECTED _OnStart : E_ActStatus
VAR_INPUT
    nAction : UINT;
END_VAR
IF GVL_IoRef.ipPlanar = 0 THEN
    _Fail(GVL_Catalog.Err_NotWired, 0);
    _OnStart := E_ActStatus.Error;
    RETURN;
END_IF
CASE nAction OF
    GVL_Catalog.PlanarSystem_ActiverLeSysteme, GVL_Catalog.PlanarSystem_DesactiverLeSysteme, GVL_Catalog.PlanarSystem_AcquitterErreur:
        _OnStart := _OnCycle(nAction);
ELSE
    _OnStart := E_ActStatus.Error;
END_CASE
END_METHOD

METHOD PROTECTED _OnCycle : E_ActStatus
VAR_INPUT
    nAction : UINT;
END_VAR
_OnCycle := E_ActStatus.Busy;
CASE nAction OF
    GVL_Catalog.PlanarSystem_ActiverLeSysteme:
        IF GVL_IoRef.ipPlanar.Activate(TRUE) THEN
            _SetResult(1, INT_TO_LREAL(_nDetected));
            _OnCycle := E_ActStatus.Done;
        END_IF
    GVL_Catalog.PlanarSystem_DesactiverLeSysteme:
        GVL_IoRef.ipPlanar.Activate(FALSE);
        IF NOT GVL_IoRef.ipPlanar.Active THEN _OnCycle := E_ActStatus.Done; END_IF
    GVL_Catalog.PlanarSystem_AcquitterErreur:
        GVL_IoRef.ipPlanar.AckError();
        IF GVL_IoRef.ipPlanar.ErrorCode = 0 THEN _OnCycle := E_ActStatus.Done; END_IF
ELSE
    _OnCycle := E_ActStatus.Error;
END_CASE
END_METHOD

METHOD PROTECTED _Publish
VAR
    i : USINT;
END_VAR
_nDetected := 0;
IF GVL_IoRef.ipPlanar = 0 THEN RETURN; END_IF
FOR i := 1 TO GVL_Const.MAX_MOVERS DO
    IF GVL_IoRef.ipPlanar.MoverDetected(i) THEN _nDetected := _nDetected + 1; END_IF
END_FOR
_stStatus.aValue[1] := SEL(GVL_IoRef.ipPlanar.Active, 0.0, 1.0);
_stStatus.aValue[2] := INT_TO_LREAL(_nDetected);
END_METHOD
END_FUNCTION_BLOCK

(* ---- FB_Press.st ---- *)
// Presse, type 40 (docs/03 § 7.1) : D axe NC de la presse, S1 AI capteur de force. Recettes déployées dans
// GVL_Active.aPressRecipe (8 segments au plus : course cible ou force cible, vitesse, fenêtres de contrôle).
// Chaque exécution enregistre la courbe force/course (1 000 points au plus) dans GVL_Hmi.aCurve.
// Hypothèses : la valeur brute de S1 est en newtons ; la position de repos est la course 0 de l'axe (la fiche
// parle d'une position nommée sans dire laquelle) ; l'axe est référencé par TwinCAT (codeur absolu) et
// alimenté tant que l'objet n'est ni en erreur ni désactivé ; une fenêtre dont les deux bornes valent 0 n'est
// pas contrôlée.
FUNCTION_BLOCK FB_Press EXTENDS FB_ObjectBase
VAR
    _pAxis : POINTER TO AXIS_REF;
    _fbPower : MC_Power;
    _fbReset : MC_Reset;
    _fbMoveAbs : MC_MoveAbsolute;
    _fbMoveVel : MC_MoveVelocity;
    _fbHalt : MC_Halt;
    _bEnable : BOOL;
    _bPowered : BOOL;
    _bAbs : BOOL;                   // commande de MC_MoveAbsolute
    _bVel : BOOL;                   // commande de MC_MoveVelocity (segment à force cible)
    _bHalt : BOOL;
    _fTarget : LREAL;
    _fVelo : LREAL;
    _fForce : LREAL;                // N, après tare
    _fForceRaw : LREAL;
    _fStroke : LREAL;               // mm
    _fForceMax : LREAL;
    _nRecipe : INT;                 // rang dans aPressRecipe
    _nRecipeNo : INT;
    _nSeg : USINT;
    _nPhase : USINT;                // 0 lancer le segment, 1 en mouvement, 2 arrêt, 3 retour repos
    _bAllOk : BOOL;
    _nCurveSlot : USINT;
    _nCurveId : UDINT;
    _fOverride : LREAL := 100.0;
    // Simulation
    _fSimStroke : LREAL;
    _fSimVel : LREAL;
    _fSimContact : LREAL;
    _fSimStiffness : LREAL := 200.0; // N/mm
    _bSimBad : BOOL;
END_VAR
VAR PERSISTENT
    _fTare : LREAL;
END_VAR

METHOD PROTECTED _OnConfigure : BOOL
IF _bNewObject THEN _fTare := 0; END_IF
_pAxis := F_AxisRef(_refCfg.nDevice);
_OnConfigure := F_SignalValid(_refCfg.aSignal[1], E_SignalKind.AI) AND (_pAxis <> 0 OR _IsSimulated());
END_METHOD

METHOD PROTECTED _IsMotion : BOOL
VAR_INPUT
    nAction : UINT;
END_VAR
_IsMotion := nAction = GVL_Catalog.Press_ExecuterRecette OR nAction = GVL_Catalog.Press_RetourRepos;
END_METHOD

METHOD PROTECTED _DefaultTimeoutMs : UDINT
VAR_INPUT
    nAction : UINT;
END_VAR
CASE nAction OF
    GVL_Catalog.Press_ExecuterRecette: _DefaultTimeoutMs := LREAL_TO_UDINT(MAX(1000.0, _refCfg.aParam[2]));
    GVL_Catalog.Press_RetourRepos: _DefaultTimeoutMs := 5000;
    GVL_Catalog.Press_TarerLaForce: _DefaultTimeoutMs := 2000;
ELSE
    _DefaultTimeoutMs := 0;
END_CASE
END_METHOD

METHOD PROTECTED _OnStart : E_ActStatus
VAR_INPUT
    nAction : UINT;
END_VAR
VAR
    k : INT;
END_VAR
CASE nAction OF
    GVL_Catalog.Press_ExecuterRecette:
        _nRecipeNo := LREAL_TO_INT(_ParamReal(1, 0));
        _nRecipe := 0;
        FOR k := 1 TO GVL_Const.MAX_PRESS_RECIPES DO
            IF GVL_Active.aPressRecipe[k].bUsed AND GVL_Active.aPressRecipe[k].nStation = _stInfo.nStation
               AND GVL_Active.aPressRecipe[k].nObject = _stInfo.nLocalId AND GVL_Active.aPressRecipe[k].nRecipeNo = _nRecipeNo THEN
                _nRecipe := k;
            END_IF
        END_FOR
        IF _nRecipe = 0 OR_ELSE GVL_Active.aPressRecipe[_nRecipe].nSegments = 0 THEN
            _Fail(GVL_Catalog.Press_Err104, INT_TO_UDINT(_nRecipeNo));
            _OnStart := E_ActStatus.Error;
            RETURN;
        END_IF
        _nSeg := 1;
        _nPhase := 0;
        _bAllOk := TRUE;
        _fForceMax := 0;
        _bSimBad := F_SimRandom() >= 0.97;          // simulation : jugement bon à 97 % (docs/03 § 7.1)
        _fSimContact := _SimContact();
        _BeginCurve();
        _OnStart := E_ActStatus.Busy;
    GVL_Catalog.Press_RetourRepos:
        _fTarget := 0;
        _fVelo := MAX(1.0, _refCfg.aParam[4] * LIMIT(1.0, _refCfg.aParam[3], 100.0) / 100.0);
        _bAbs := FALSE;
        _nPhase := 3;
        _OnStart := E_ActStatus.Busy;
    GVL_Catalog.Press_TarerLaForce:
        _fTare := _fForceRaw;
        _OnStart := E_ActStatus.Done;
    GVL_Catalog.Press_LireForceEtCourse:
        _SetResult(1, _fForce);
        _SetResult(2, _fStroke);
        _OnStart := E_ActStatus.Done;
ELSE
    _OnStart := E_ActStatus.Error;
END_CASE
END_METHOD

METHOD PROTECTED _OnCycle : E_ActStatus
VAR_INPUT
    nAction : UINT;
END_VAR
VAR
    s : REFERENCE TO ST_PressSegment;
    bReached : BOOL;
END_VAR
_OnCycle := E_ActStatus.Busy;
// Force maximale de sécurité : arrêt immédiat, défaut (erreur 100)
IF _fForce > MAX(1.0, _refCfg.aParam[1]) THEN
    _StopMotion();
    _Fail(GVL_Catalog.Press_Err100, LREAL_TO_UDINT(_fForce));
    _OnCycle := E_ActStatus.Error;
    RETURN;
END_IF
IF _nPhase = 3 THEN
    // Retour repos
    IF NOT _bAbs THEN _bAbs := TRUE; RETURN; END_IF
    IF _MoveDone() THEN _bAbs := FALSE; _nPhase := 0; _OnCycle := E_ActStatus.Done; END_IF
    IF _MoveError() THEN _bAbs := FALSE; _Fail(GVL_Catalog.Press_Err101, 0); _OnCycle := E_ActStatus.Error; END_IF
    RETURN;
END_IF
_RecordPoint();
_fForceMax := MAX(_fForceMax, _fForce);
s REF= GVL_Active.aPressRecipe[_nRecipe].aSeg[_nSeg];
CASE _nPhase OF
    0:  // lancer le segment : course cible en position, force cible en vitesse jusqu'à la force
        _fVelo := MAX(0.1, _refCfg.aParam[4] * LIMIT(1.0, s.fSpeedPct, 100.0) / 100.0);
        IF s.eTarget = 0 THEN
            _fTarget := s.fTarget;
            _bAbs := TRUE;
        ELSE
            _bVel := TRUE;
        END_IF
        _nPhase := 1;
    1:
        IF s.eTarget = 0 THEN
            bReached := _MoveDone();
        ELSE
            bReached := _fForce >= s.fTarget;
        END_IF
        IF _MoveError() THEN
            _StopMotion();
            _Fail(GVL_Catalog.Press_Err101, _nSeg);
            _OnCycle := E_ActStatus.Error;
            RETURN;
        END_IF
        IF bReached THEN
            _bAbs := FALSE;
            IF _bVel THEN _bVel := FALSE; _bHalt := TRUE; _nPhase := 2; ELSE _EndSegment(); END_IF
        ELSIF s.eTarget = 1 AND _fStroke >= _MaxStroke(s) THEN
            _StopMotion();                                  // force non atteinte avant la course maximale
            _Fail(GVL_Catalog.Press_Err103, _nSeg);
            _OnCycle := E_ActStatus.Error;
            RETURN;
        END_IF
    2:
        IF _HaltDone() THEN
            _bHalt := FALSE;
            _EndSegment();
        END_IF
END_CASE
IF _nSeg > GVL_Active.aPressRecipe[_nRecipe].nSegments THEN
    _EndCurve();
    _SetJudgement(1, SEL(_bAllOk, E_Judgement.Nok, E_Judgement.Ok));
    _SetResult(2, _fForce);
    _SetResult(3, _fStroke);
    _SetResult(4, _fForceMax);
    _OnCycle := E_ActStatus.Done;
END_IF
END_METHOD

// Fin d'un segment : contrôle des fenêtres de force et de course
METHOD PRIVATE _EndSegment
VAR
    s : REFERENCE TO ST_PressSegment;
END_VAR
s REF= GVL_Active.aPressRecipe[_nRecipe].aSeg[_nSeg];
IF NOT (s.fForceMin = 0 AND s.fForceMax = 0) AND (_fForce < s.fForceMin OR _fForce > s.fForceMax) THEN _bAllOk := FALSE; END_IF
IF NOT (s.fStrokeMin = 0 AND s.fStrokeMax = 0) AND (_fStroke < s.fStrokeMin OR _fStroke > s.fStrokeMax) THEN _bAllOk := FALSE; END_IF
_nSeg := _nSeg + 1;
_nPhase := 0;
END_METHOD

// Course maximale d'un segment à force cible : borne haute de sa fenêtre de course, sinon 200 mm
METHOD PRIVATE _MaxStroke : LREAL
VAR_INPUT
    s : REFERENCE TO ST_PressSegment;
END_VAR
IF s.fStrokeMax > 0 THEN _MaxStroke := s.fStrokeMax; ELSE _MaxStroke := 200.0; END_IF
END_METHOD

METHOD PROTECTED _OnAbort
VAR_INPUT
    nAction : UINT;
END_VAR
_StopMotion();
_EndCurve();
END_METHOD

METHOD PROTECTED _SafeState
_StopMotion();
END_METHOD

METHOD PRIVATE _StopMotion
_bAbs := FALSE;
_bVel := FALSE;
_bHalt := _bPowered AND NOT _IsSimulated();
_fSimVel := 0;
END_METHOD

METHOD PRIVATE _MoveDone : BOOL
IF _IsSimulated() THEN
    _MoveDone := ABS(_fSimStroke - _fTarget) < 0.001;
ELSE
    _MoveDone := _fbMoveAbs.Done;
END_IF
END_METHOD

METHOD PRIVATE _MoveError : BOOL
_MoveError := NOT _IsSimulated() AND (_fbMoveAbs.Error OR _fbMoveVel.Error OR _fbPower.Error);
END_METHOD

METHOD PRIVATE _HaltDone : BOOL
_HaltDone := _IsSimulated() OR _fbHalt.Done OR _fbHalt.Error;
END_METHOD

// ---------- courbe force/course (docs/05 § 9)

METHOD PRIVATE _BeginCurve
_nCurveSlot := GVL_Curves.nNextSlot;
GVL_Curves.nNextSlot := GVL_Curves.nNextSlot MOD GVL_Const.CURVE_BUFFER + 1;
_nCurveId := GVL_Curves.nNextCurveId;
GVL_Curves.nNextCurveId := GVL_Curves.nNextCurveId + 1;
GVL_Hmi.aCurve[_nCurveSlot].nCurveId := 0;          // invalide tant qu'elle s'écrit
GVL_Hmi.aCurve[_nCurveSlot].nPoints := 0;
IF _stInfo.nStation <= GVL_Const.MAX_STATIONS THEN
    GVL_Curves.aLastCurveId[_stInfo.nStation] := _nCurveId;
    GVL_Curves.aLastCurveTime[_stInfo.nStation] := F_NowUtc();
END_IF
END_METHOD

METHOD PRIVATE _RecordPoint
VAR
    c : REFERENCE TO ST_PressCurve;
END_VAR
IF _nCurveSlot = 0 THEN RETURN; END_IF
c REF= GVL_Hmi.aCurve[_nCurveSlot];
IF c.nPoints < GVL_Const.CURVE_POINTS THEN
    c.nPoints := c.nPoints + 1;
    c.aStroke[c.nPoints] := LREAL_TO_REAL(_fStroke);
    c.aForce[c.nPoints] := LREAL_TO_REAL(_fForce);
END_IF
END_METHOD

METHOD PRIVATE _EndCurve
IF _nCurveSlot = 0 THEN RETURN; END_IF
GVL_Hmi.aCurve[_nCurveSlot].nCurveId := _nCurveId;
_nCurveSlot := 0;
END_METHOD

// ---------- matériel et simulation

METHOD PROTECTED _ApplyOverride
VAR_INPUT
    fPercent : LREAL;
END_VAR
_fOverride := fPercent;
END_METHOD

METHOD PROTECTED _ReadHw
_fForceRaw := INT_TO_LREAL(F_ReadAI(_refCfg.aSignal[1]));
_fForce := _fForceRaw - _fTare;
IF _pAxis <> 0 THEN _fStroke := _pAxis^.NcToPlc.ActPos; END_IF
END_METHOD

METHOD PROTECTED _WriteHw
IF _IsSimulated() OR _pAxis = 0 THEN RETURN; END_IF
_bEnable := _eState <> E_ObjState.Error AND _eState <> E_ObjState.Disabled;
_fbPower(Axis := _pAxis^, Enable := _bEnable, Enable_Positive := _bEnable, Enable_Negative := _bEnable, Override := _fOverride);
_bPowered := _fbPower.Status;
_fbMoveAbs(Axis := _pAxis^, Execute := _bAbs, Position := _fTarget, Velocity := _fVelo);
_fbMoveVel(Axis := _pAxis^, Execute := _bVel, Velocity := _fVelo, Direction := MC_Positive_Direction);
_fbHalt(Axis := _pAxis^, Execute := _bHalt);
_fbReset(Axis := _pAxis^, Execute := _eState = E_ObjState.Error AND _fbPower.Error);
END_METHOD

// Simulation : course intégrée à la vitesse commandée, force nulle avant le contact puis raideur constante
METHOD PROTECTED _Simulate
VAR
    fStep : LREAL;
END_VAR
_bPowered := TRUE;
fStep := _fVelo * F_CycleMs() / 1000.0 * _fOverride / 100.0;
IF _bAbs THEN
    IF _fSimStroke < _fTarget THEN _fSimStroke := MIN(_fTarget, _fSimStroke + fStep); ELSE _fSimStroke := MAX(_fTarget, _fSimStroke - fStep); END_IF
ELSIF _bVel THEN
    _fSimStroke := _fSimStroke + fStep;
END_IF
_fStroke := _fSimStroke;
_fForceRaw := MAX(0.0, (_fSimStroke - _fSimContact) * _fSimStiffness) + _fTare;
IF _Forced(1) THEN _fForceRaw := _ForcedValue(1) + _fTare; END_IF
_fForce := _fForceRaw - _fTare;
END_METHOD

// Course du contact simulé : au milieu de la fenêtre de force du dernier segment, décalée si le tirage est mauvais
METHOD PRIVATE _SimContact : LREAL
VAR
    s : REFERENCE TO ST_PressSegment;
    fWanted : LREAL;
END_VAR
s REF= GVL_Active.aPressRecipe[_nRecipe].aSeg[GVL_Active.aPressRecipe[_nRecipe].nSegments];
IF s.eTarget = 0 THEN
    IF s.fForceMax > 0 THEN fWanted := (s.fForceMin + s.fForceMax) / 2.0; ELSE fWanted := 500.0; END_IF
    _SimContact := s.fTarget - fWanted / _fSimStiffness;
    IF _bSimBad THEN _SimContact := _SimContact - 2.0 * MAX(1.0, (s.fForceMax - s.fForceMin)) / _fSimStiffness; END_IF
ELSE
    _SimContact := MAX(1.0, s.fStrokeMin + (s.fStrokeMax - s.fStrokeMin) / 2.0 - s.fTarget / _fSimStiffness);
    IF _bSimBad THEN _SimContact := _SimContact + MAX(1.0, s.fStrokeMax - s.fStrokeMin); END_IF
END_IF
END_METHOD

METHOD PROTECTED _Publish
_stStatus.aValue[1] := _fForce;
_stStatus.aValue[2] := _fStroke;
_stStatus.aValue[3] := INT_TO_LREAL(_nRecipeNo);
END_METHOD
END_FUNCTION_BLOCK

(* ---- FB_Safety.st ---- *)
// Sécurités, type 51 (docs/03 § 8.2) : lit les retours des circuits (1 = OK), ne pilote rien, aucun contournement.
// Un circuit ouvert met l'objet en erreur 100 (défaut machine ou de station selon son emplacement) ; un circuit qui
// demande un acquittement reste « à acquitter » (erreur 102) jusqu'à l'action Acquitter ou l'Ack de l'objet.
FUNCTION_BLOCK FB_Safety EXTENDS FB_ObjectBase IMPLEMENTS I_SafetyCircuits
VAR
    _aRaw : ARRAY[1..8] OF BOOL;
    _aOk : ARRAY[1..8] OF BOOL;         // filtré
    _aFilter : ARRAY[1..8] OF LREAL;
    _aToAck : ARRAY[1..8] OF BOOL;
    _aUsed : ARRAY[1..8] OF BOOL;
    _nCircuit : INT;
END_VAR

METHOD PROTECTED _OnConfigure : BOOL
VAR
    i : USINT;
END_VAR
FOR i := 1 TO 8 DO
    _aUsed[i] := F_SignalValid(_refCfg.aSignal[i], E_SignalKind.DI);
    _aOk[i] := TRUE;
    _aRaw[i] := TRUE;
    _aToAck[i] := FALSE;
END_FOR
_OnConfigure := TRUE;
END_METHOD

PROPERTY AllOk : BOOL
GET
VAR
    i : INT;
END_VAR
AllOk := TRUE;
FOR i := 1 TO 8 DO
    IF _aUsed[i] AND (NOT _aOk[i] OR _aToAck[i]) THEN AllOk := FALSE; END_IF
END_FOR
END_GET
END_PROPERTY

METHOD PRIVATE _CircuitOk : BOOL
VAR_INPUT
    nCircuit : INT;              // 0 = tous
END_VAR
VAR
    i : INT;
END_VAR
_CircuitOk := TRUE;
FOR i := 1 TO 8 DO
    IF _aUsed[i] AND (nCircuit = 0 OR nCircuit = i) AND (NOT _aOk[i] OR _aToAck[i]) THEN _CircuitOk := FALSE; END_IF
END_FOR
END_METHOD

METHOD PRIVATE _AckCircuits : BOOL
VAR_INPUT
    nCircuit : INT;
END_VAR
VAR
    i : INT;
END_VAR
_AckCircuits := TRUE;
FOR i := 1 TO 8 DO
    IF (nCircuit = 0 OR nCircuit = i) AND _aToAck[i] THEN
        IF _aOk[i] THEN _aToAck[i] := FALSE; ELSE _AckCircuits := FALSE; END_IF
    END_IF
END_FOR
END_METHOD

METHOD PROTECTED _OnStart : E_ActStatus
VAR_INPUT
    nAction : UINT;
END_VAR
_nCircuit := LIMIT(0, LREAL_TO_INT(_ParamReal(1, 0.0)), 8);
CASE nAction OF
    GVL_Catalog.Safety_LireEtat:
        _SetResult(1, BOOL_TO_LREAL(_CircuitOk(_nCircuit)));
        _OnStart := E_ActStatus.Done;
    GVL_Catalog.Safety_Acquitter, GVL_Catalog.Safety_AttendreOK:
        _OnStart := _OnCycle(nAction);
ELSE
    _OnStart := E_ActStatus.Error;
END_CASE
END_METHOD

METHOD PROTECTED _OnCycle : E_ActStatus
VAR_INPUT
    nAction : UINT;
END_VAR
IF nAction = GVL_Catalog.Safety_Acquitter THEN
    IF _AckCircuits(_nCircuit) THEN _OnCycle := E_ActStatus.Done; ELSE _OnCycle := E_ActStatus.Busy; END_IF
ELSIF _CircuitOk(_nCircuit) THEN
    _OnCycle := E_ActStatus.Done;
ELSE
    _OnCycle := E_ActStatus.Busy;
END_IF
END_METHOD

METHOD PROTECTED _OnAck : BOOL
_OnAck := _AckCircuits(0) AND _CircuitOk(0);
END_METHOD

METHOD PROTECTED _Monitor
VAR
    i : INT;
END_VAR
FOR i := 1 TO 8 DO
    IF _aUsed[i] THEN
        IF _aRaw[i] = _aOk[i] THEN
            _aFilter[i] := 0;
        ELSE
            _aFilter[i] := _aFilter[i] + F_CycleMs();
            IF _aFilter[i] >= _refCfg.aParam[17] THEN
                _aOk[i] := _aRaw[i];
                _aFilter[i] := 0;
                IF NOT _aOk[i] AND _refCfg.aParam[8 + i] = 1 THEN _aToAck[i] := TRUE; END_IF
            END_IF
        END_IF
        IF NOT _aOk[i] AND _eState <> E_ObjState.Error THEN
            _Fail(GVL_Catalog.Safety_Err100, INT_TO_UDINT(i));            // circuit ouvert
        ELSIF _aOk[i] AND _aToAck[i] AND _eState <> E_ObjState.Error THEN
            _Fail(GVL_Catalog.Safety_Err102, INT_TO_UDINT(i));            // acquittement requis
        END_IF
    END_IF
END_FOR
END_METHOD

METHOD PROTECTED _ReadHw
VAR
    i : USINT;
END_VAR
FOR i := 1 TO 8 DO
    IF _aUsed[i] THEN _aRaw[i] := F_ReadDI(_refCfg.aSignal[i]); END_IF
END_FOR
END_METHOD

METHOD PROTECTED _Simulate
VAR
    i : USINT;
END_VAR
FOR i := 1 TO 8 DO
    IF _Forced(i) THEN _aRaw[i] := _ForcedValue(i) >= 0.5; ELSE _aRaw[i] := TRUE; END_IF
END_FOR
END_METHOD

METHOD PROTECTED _Publish
VAR
    i : INT;
    nOk : DWORD;
    nAck : DWORD;
END_VAR
FOR i := 1 TO 8 DO
    IF _aUsed[i] AND _aOk[i] THEN nOk := nOk OR SHL(DWORD#1, i - 1); END_IF
    IF _aToAck[i] THEN nAck := nAck OR SHL(DWORD#1, i - 1); END_IF
END_FOR
_stStatus.aValue[1] := DWORD_TO_LREAL(nOk);
_stStatus.aValue[2] := DWORD_TO_LREAL(nAck);
END_METHOD
END_FUNCTION_BLOCK

(* ---- FB_Scale.st ---- *)
// Pesage, type 33 (docs/03 § 6.4), mode analogique : S1 AI mesure. Le mode réseau n'est pas encore écrit.
// Hypothèses : la valeur brute est en dixièmes de l'unité P1 (g ou mg) ; la mesure est stable quand l'écart
// entre la plus grande et la plus petite des 10 dernières valeurs ne dépasse pas 0,5 unité ; tolérance basse
// P3 négative ou positive, prise en valeur absolue sous la valeur nominale P4.
FUNCTION_BLOCK FB_Scale EXTENDS FB_ObjectBase
VAR
    _fGross : LREAL;
    _fValue : LREAL;
    _bOverload : BOOL;
    _aWin : ARRAY[1..10] OF LREAL;
    _nWin : INT;
    _nNext : INT := 1;
    _bStable : BOOL;
    _fStabMs : LREAL;
    _nWanted : INT;
    _nTaken : INT;
    _fSum : LREAL;
END_VAR
VAR PERSISTENT
    _fTare : LREAL;
END_VAR

METHOD PROTECTED _OnConfigure : BOOL
IF _bNewObject THEN _fTare := 0; END_IF
_nWin := 0;
_nNext := 1;
_OnConfigure := F_SignalValid(_refCfg.aSignal[1], E_SignalKind.AI);
END_METHOD

METHOD PROTECTED _OnStart : E_ActStatus
VAR_INPUT
    nAction : UINT;
END_VAR
CASE nAction OF
    GVL_Catalog.Scale_Tarer, GVL_Catalog.Scale_Mesurer:
        _nWanted := LIMIT(1, LREAL_TO_INT(_ParamReal(1, _refCfg.aParam[5])), 1000);
        _nTaken := 0;
        _fSum := 0;
        _fStabMs := 0;
        _OnStart := E_ActStatus.Busy;
    GVL_Catalog.Scale_LireValeurCourante:
        _SetResult(1, _fValue);
        _SetResult(2, SEL(_bStable, 0.0, 1.0));
        _OnStart := E_ActStatus.Done;
ELSE
    _OnStart := E_ActStatus.Error;
END_CASE
END_METHOD

METHOD PROTECTED _OnCycle : E_ActStatus
VAR_INPUT
    nAction : UINT;
END_VAR
VAR
    fMean : LREAL;
    fLow : LREAL;
END_VAR
_OnCycle := E_ActStatus.Busy;
IF _bOverload THEN
    _Fail(GVL_Catalog.Scale_Err101, 0);
    _OnCycle := E_ActStatus.Error;
    RETURN;
END_IF
_fStabMs := _fStabMs + F_CycleMs();
IF _fStabMs < MAX(0.0, _refCfg.aParam[6]) THEN RETURN; END_IF
IF NOT _bStable THEN
    // Pas stable deux fois le temps de stabilisation après son début : erreur 100
    IF _fStabMs >= 2.0 * MAX(100.0, _refCfg.aParam[6]) THEN
        _Fail(GVL_Catalog.Scale_Err100, 0);
        _OnCycle := E_ActStatus.Error;
    END_IF
    RETURN;
END_IF
IF nAction = GVL_Catalog.Scale_Tarer THEN
    _fTare := _fGross;
    _OnCycle := E_ActStatus.Done;
    RETURN;
END_IF
_fSum := _fSum + _fValue;
_nTaken := _nTaken + 1;
IF _nTaken < _nWanted THEN RETURN; END_IF
fMean := _fSum / INT_TO_LREAL(_nTaken);
_SetResult(1, fMean);
fLow := _refCfg.aParam[4] - ABS(_refCfg.aParam[3]);
IF _refCfg.aParam[2] = 0 AND _refCfg.aParam[3] = 0 THEN
    _SetJudgement(2, E_Judgement.Ok);           // pas de tolérance : pas de jugement
ELSIF fMean > _refCfg.aParam[4] + ABS(_refCfg.aParam[2]) THEN
    _SetJudgement(2, E_Judgement.High);
ELSIF fMean < fLow THEN
    _SetJudgement(2, E_Judgement.Low);
ELSE
    _SetJudgement(2, E_Judgement.Ok);
END_IF
_OnCycle := E_ActStatus.Done;
END_METHOD

METHOD PROTECTED _ReadHw
VAR
    nRaw : INT;
END_VAR
nRaw := F_ReadAI(_refCfg.aSignal[1]);
_bOverload := nRaw = 32767;
_Sample(INT_TO_LREAL(nRaw) * 0.1);
END_METHOD

// Simulation : valeur nominale P4 (plus la tare) avec un bruit de ±0,1 unité
METHOD PROTECTED _Simulate
VAR
    fGross : LREAL;
END_VAR
fGross := _refCfg.aParam[4] + _fTare + (F_SimRandom() - 0.5) * 0.2;
IF _Forced(1) THEN fGross := _ForcedValue(1) + _fTare; END_IF       // valeur forcée nette, en unité
_bOverload := FALSE;
_Sample(fGross);
END_METHOD

METHOD PRIVATE _Sample
VAR_INPUT
    fGross : LREAL;
END_VAR
VAR
    i : INT;
    fMin : LREAL := 1.0E38;
    fMax : LREAL := -1.0E38;
END_VAR
_fGross := fGross;
_fValue := fGross - _fTare;
_aWin[_nNext] := fGross;
_nNext := _nNext MOD 10 + 1;
_nWin := MIN(_nWin + 1, 10);
FOR i := 1 TO _nWin DO
    fMin := MIN(fMin, _aWin[i]);
    fMax := MAX(fMax, _aWin[i]);
END_FOR
_bStable := _nWin = 10 AND fMax - fMin <= 0.5;
END_METHOD

METHOD PROTECTED _Publish
_stStatus.aValue[1] := _fValue;
_stStatus.aValue[2] := SEL(_bStable, 0.0, 1.0);
END_METHOD
END_FUNCTION_BLOCK

(* ---- FB_Timer.st ---- *)
// Temporisation, type 52 (docs/03 § 8.3)
FUNCTION_BLOCK FB_Timer EXTENDS FB_ObjectBase
VAR
    _fDurationMs : LREAL;
    _fElapsed : LREAL;
END_VAR

METHOD PROTECTED _OnStart : E_ActStatus
VAR_INPUT
    nAction : UINT;
END_VAR
IF nAction = GVL_Catalog.Timer_Attendre THEN
    _fDurationMs := MAX(0.0, _ParamReal(1, _refCfg.aParam[1]));
    _fElapsed := 0;
    _OnStart := _OnCycle(nAction);
ELSE
    _OnStart := E_ActStatus.Error;
END_IF
END_METHOD

METHOD PROTECTED _OnCycle : E_ActStatus
VAR_INPUT
    nAction : UINT;
END_VAR
_fElapsed := _fElapsed + F_CycleMs();
IF _fElapsed >= _fDurationMs THEN _OnCycle := E_ActStatus.Done; ELSE _OnCycle := E_ActStatus.Busy; END_IF
END_METHOD

METHOD PROTECTED _DefaultTimeoutMs : UDINT
VAR_INPUT
    nAction : UINT;
END_VAR
_DefaultTimeoutMs := 0;             // aucun timeout (docs/03 § 8.3)
END_METHOD

METHOD PROTECTED _Publish
IF _eState = E_ObjState.Busy AND _fDurationMs > 0 THEN
    _stStatus.fProgress := LREAL_TO_REAL(MIN(1.0, _fElapsed / _fDurationMs));
END_IF
END_METHOD
END_FUNCTION_BLOCK

(* ---- FB_VacuumBlow.st ---- *)
// Aspiration et soufflage, type 20 (docs/03 § 5.1).
// Capteur de vide : S3 pressostat (DI) ou S4 analogique. Hypothèse (à confirmer) : l'entrée analogique donne le vide
// en dixièmes de kPa (valeur brute ÷ 10).
FUNCTION_BLOCK FB_VacuumBlow EXTENDS FB_ObjectBase
VAR
    _bSuck : BOOL;
    _bBlow : BOOL;
    _bHasBlow : BOOL;
    _bDigital : BOOL;               // pressostat S3
    _bAnalog : BOOL;                // capteur S4
    _fVacuum : LREAL;               // kPa (négatif), ou 0/1 pour le pressostat
    _bPresent : BOOL;
    _bEmptyNozzle : BOOL;           // vide sous le seuil « buse vide »
    _bHolding : BOOL;               // pièce prise : une perte de vide est une erreur 101
    _bWaitVacuum : BOOL;
    _fBlowMs : LREAL;
    _fElapsed : LREAL;
    _fSimVacuum : LREAL;
END_VAR

METHOD PROTECTED _OnConfigure : BOOL
_bHasBlow := F_SignalValid(_refCfg.aSignal[2], E_SignalKind.DO);
_bDigital := F_SignalValid(_refCfg.aSignal[3], E_SignalKind.DI);
_bAnalog := F_SignalValid(_refCfg.aSignal[4], E_SignalKind.AI);
_bHolding := FALSE;
_OnConfigure := F_SignalValid(_refCfg.aSignal[1], E_SignalKind.DO) AND (_bDigital OR _bAnalog);
END_METHOD

METHOD PROTECTED _DefaultTimeoutMs : UDINT
VAR_INPUT
    nAction : UINT;
END_VAR
IF nAction = GVL_Catalog.VacuumBlow_Souffler THEN
    _DefaultTimeoutMs := LREAL_TO_UDINT(_ParamReal(1, _refCfg.aParam[3])) + 500;
ELSE
    _DefaultTimeoutMs := SUPER^._DefaultTimeoutMs(nAction);
END_IF
END_METHOD

METHOD PROTECTED _OnStart : E_ActStatus
VAR_INPUT
    nAction : UINT;
END_VAR
_fElapsed := 0;
CASE nAction OF
    GVL_Catalog.VacuumBlow_Aspirer:
        _bBlow := FALSE;
        _bSuck := TRUE;
        _bWaitVacuum := _ParamReal(1, 1.0) >= 0.5;
        IF NOT _bWaitVacuum THEN
            _SetResult(1, BOOL_TO_LREAL(_bPresent));
            _OnStart := E_ActStatus.Done;
        ELSE
            _OnStart := E_ActStatus.Busy;
        END_IF
    GVL_Catalog.VacuumBlow_Souffler:
        _bSuck := FALSE;
        _bHolding := FALSE;
        _fBlowMs := MAX(_ParamReal(1, _refCfg.aParam[3]), 0.0);
        _bBlow := _bHasBlow;
        _OnStart := E_ActStatus.Busy;
    GVL_Catalog.VacuumBlow_Couper:
        _bSuck := FALSE;
        _bBlow := FALSE;
        _bHolding := FALSE;
        _OnStart := E_ActStatus.Done;
    GVL_Catalog.VacuumBlow_VerifierPresencePiece:
        _SetResult(1, BOOL_TO_LREAL(_bPresent));
        _OnStart := E_ActStatus.Done;
ELSE
    _OnStart := E_ActStatus.Error;
END_CASE
END_METHOD

METHOD PROTECTED _OnCycle : E_ActStatus
VAR_INPUT
    nAction : UINT;
END_VAR
_fElapsed := _fElapsed + F_CycleMs();
CASE nAction OF
    GVL_Catalog.VacuumBlow_Aspirer:
        IF _bPresent THEN
            _bHolding := TRUE;
            _SetResult(1, 1.0);
            _OnCycle := E_ActStatus.Done;
        ELSIF _nTimeoutMs > 0 AND _fElapsed + F_CycleMs() >= UDINT_TO_LREAL(_nTimeoutMs) THEN
            _Fail(GVL_Catalog.VacuumBlow_Err100, 0);        // vide non atteint, avant le timeout générique
            _OnCycle := E_ActStatus.Error;
        ELSE
            _OnCycle := E_ActStatus.Busy;
        END_IF
    GVL_Catalog.VacuumBlow_Souffler:
        IF _fElapsed >= _fBlowMs THEN
            _bBlow := FALSE;
            _OnCycle := E_ActStatus.Done;
        ELSE
            _OnCycle := E_ActStatus.Busy;
        END_IF
ELSE
    _OnCycle := E_ActStatus.Done;
END_CASE
END_METHOD

METHOD PROTECTED _OnAbort
VAR_INPUT
    nAction : UINT;
END_VAR
_bBlow := FALSE;
END_METHOD

METHOD PROTECTED _SafeState
_bBlow := FALSE;
IF _refCfg.aParam[4] = 0 THEN
    _bSuck := FALSE;                // tout couper
    _bHolding := FALSE;
END_IF                              // 1 : maintenir l'aspiration
END_METHOD

METHOD PROTECTED _Monitor
IF _bAnalog AND _refCfg.aParam[1] >= _refCfg.aParam[2] THEN
    IF _eState <> E_ObjState.Error THEN _Fail(GVL_Catalog.VacuumBlow_Err102, 0); END_IF
    RETURN;
END_IF
IF _bHolding AND _bSuck AND NOT _bPresent AND _eState <> E_ObjState.Error THEN
    _bHolding := FALSE;
    _Fail(GVL_Catalog.VacuumBlow_Err101, 0);       // pièce tombée
END_IF
END_METHOD

METHOD PROTECTED _ReadHw
IF _bDigital THEN
    _bPresent := F_ReadDI(_refCfg.aSignal[3]);
    _fVacuum := BOOL_TO_LREAL(_bPresent);
ELSE
    _fVacuum := INT_TO_LREAL(F_ReadAI(_refCfg.aSignal[4])) / 10.0;
    _Evaluate();
END_IF
END_METHOD

METHOD PROTECTED _Simulate
VAR
    fStep : LREAL;
END_VAR
// Vide simulé : −70 kPa en 80 ms quand on aspire, retour à 0 sinon
fStep := 70.0 * F_CycleMs() / 80.0;
IF _bSuck THEN _fSimVacuum := MAX(-70.0, _fSimVacuum - fStep); ELSE _fSimVacuum := MIN(0.0, _fSimVacuum + fStep); END_IF
IF _Forced(4) THEN _fSimVacuum := _ForcedValue(4); END_IF
IF _bDigital THEN
    _bPresent := _fSimVacuum <= -60.0;
    IF _Forced(3) THEN _bPresent := _ForcedValue(3) >= 0.5; END_IF
    _fVacuum := BOOL_TO_LREAL(_bPresent);
ELSE
    _fVacuum := _fSimVacuum;
    _Evaluate();
END_IF
END_METHOD

METHOD PRIVATE _Evaluate
// Hystérésis entre P1 (pièce présente, −60 kPa) et P2 (buse vide, −52 kPa)
IF _fVacuum <= _refCfg.aParam[1] THEN
    _bPresent := TRUE;
ELSIF _fVacuum >= _refCfg.aParam[2] THEN
    _bPresent := FALSE;
END_IF
_bEmptyNozzle := _fVacuum >= _refCfg.aParam[2];
END_METHOD

METHOD PROTECTED _WriteHw
F_WriteDO(_refCfg.aSignal[1], _bSuck AND NOT _bBlow);     // jamais les deux ensemble
IF _bHasBlow THEN F_WriteDO(_refCfg.aSignal[2], _bBlow AND NOT _bSuck); END_IF
END_METHOD

METHOD PROTECTED _Publish
_stStatus.aValue[1] := BOOL_TO_LREAL(_bSuck);
_stStatus.aValue[2] := BOOL_TO_LREAL(_bBlow);
_stStatus.aValue[3] := _fVacuum;
_stStatus.aValue[4] := BOOL_TO_LREAL(_bPresent);
END_METHOD
END_FUNCTION_BLOCK
